(* IEC 61131-3 sources: BODAS-HelloWorld/st/bodas_rc18_12_40/plc_logic/application/02_easyconfig/dsm_easyconfig/structure, 701 files *)

(* ---- dfc_bds_nodeb0x8000-DFC_bds_NoDeb0x8000.st ---- *)
(* --- Interface --- *)
{attribute 'external_name' := 'cmp_rts_DFC_bds_NoDeb0x8000'}
TYPE DFC_bds_NoDeb0x8000 : STRUCT
		DTC            : UDINT := 16#800000;
		DFCid          : UINT  := 721;
		debounceMethod : USINT := NO_DEBOUNCE;
	END_STRUCT
END_TYPE

(* ---- dfc_bds_nodeb0x8001-DFC_bds_NoDeb0x8001.st ---- *)
(* --- Interface --- *)
{attribute 'external_name' := 'cmp_rts_DFC_bds_NoDeb0x8001'}
TYPE DFC_bds_NoDeb0x8001 : STRUCT
		DTC            : UDINT := 16#800100;
		DFCid          : UINT  := 722;
		debounceMethod : USINT := NO_DEBOUNCE;
	END_STRUCT
END_TYPE

(* ---- dfc_bds_nodeb0x8002-DFC_bds_NoDeb0x8002.st ---- *)
(* --- Interface --- *)
{attribute 'external_name' := 'cmp_rts_DFC_bds_NoDeb0x8002'}
TYPE DFC_bds_NoDeb0x8002 : STRUCT
		DTC            : UDINT := 16#800200;
		DFCid          : UINT  := 723;
		debounceMethod : USINT := NO_DEBOUNCE;
	END_STRUCT
END_TYPE

(* ---- dfc_bds_nodeb0x8003-DFC_bds_NoDeb0x8003.st ---- *)
(* --- Interface --- *)
{attribute 'external_name' := 'cmp_rts_DFC_bds_NoDeb0x8003'}
TYPE DFC_bds_NoDeb0x8003 : STRUCT
		DTC            : UDINT := 16#800300;
		DFCid          : UINT  := 724;
		debounceMethod : USINT := NO_DEBOUNCE;
	END_STRUCT
END_TYPE

(* ---- dfc_bds_nodeb0x8004-DFC_bds_NoDeb0x8004.st ---- *)
(* --- Interface --- *)
{attribute 'external_name' := 'cmp_rts_DFC_bds_NoDeb0x8004'}
TYPE DFC_bds_NoDeb0x8004 : STRUCT
		DTC            : UDINT := 16#800400;
		DFCid          : UINT  := 725;
		debounceMethod : USINT := NO_DEBOUNCE;
	END_STRUCT
END_TYPE

(* ---- dfc_bds_nodeb0x8005-DFC_bds_NoDeb0x8005.st ---- *)
(* --- Interface --- *)
{attribute 'external_name' := 'cmp_rts_DFC_bds_NoDeb0x8005'}
TYPE DFC_bds_NoDeb0x8005 : STRUCT
		DTC            : UDINT := 16#800500;
		DFCid          : UINT  := 726;
		debounceMethod : USINT := NO_DEBOUNCE;
	END_STRUCT
END_TYPE

(* ---- dfc_bds_nodeb0x8006-DFC_bds_NoDeb0x8006.st ---- *)
(* --- Interface --- *)
{attribute 'external_name' := 'cmp_rts_DFC_bds_NoDeb0x8006'}
TYPE DFC_bds_NoDeb0x8006 : STRUCT
		DTC            : UDINT := 16#800600;
		DFCid          : UINT  := 727;
		debounceMethod : USINT := NO_DEBOUNCE;
	END_STRUCT
END_TYPE

(* ---- dfc_bds_nodeb0x8007-DFC_bds_NoDeb0x8007.st ---- *)
(* --- Interface --- *)
{attribute 'external_name' := 'cmp_rts_DFC_bds_NoDeb0x8007'}
TYPE DFC_bds_NoDeb0x8007 : STRUCT
		DTC            : UDINT := 16#800700;
		DFCid          : UINT  := 728;
		debounceMethod : USINT := NO_DEBOUNCE;
	END_STRUCT
END_TYPE

(* ---- dfc_bds_nodeb0x8008-DFC_bds_NoDeb0x8008.st ---- *)
(* --- Interface --- *)
{attribute 'external_name' := 'cmp_rts_DFC_bds_NoDeb0x8008'}
TYPE DFC_bds_NoDeb0x8008 : STRUCT
		DTC            : UDINT := 16#800800;
		DFCid          : UINT  := 729;
		debounceMethod : USINT := NO_DEBOUNCE;
	END_STRUCT
END_TYPE

(* ---- dfc_bds_nodeb0x8009-DFC_bds_NoDeb0x8009.st ---- *)
(* --- Interface --- *)
{attribute 'external_name' := 'cmp_rts_DFC_bds_NoDeb0x8009'}
TYPE DFC_bds_NoDeb0x8009 : STRUCT
		DTC            : UDINT := 16#800900;
		DFCid          : UINT  := 730;
		debounceMethod : USINT := NO_DEBOUNCE;
	END_STRUCT
END_TYPE

(* ---- dfc_bds_nodeb0x800a-DFC_bds_NoDeb0x800a.st ---- *)
(* --- Interface --- *)
{attribute 'external_name' := 'cmp_rts_DFC_bds_NoDeb0x800a'}
TYPE DFC_bds_NoDeb0x800a : STRUCT
		DTC            : UDINT := 16#800A00;
		DFCid          : UINT  := 731;
		debounceMethod : USINT := NO_DEBOUNCE;
	END_STRUCT
END_TYPE

(* ---- dfc_bds_nodeb0x800b-DFC_bds_NoDeb0x800b.st ---- *)
(* --- Interface --- *)
{attribute 'external_name' := 'cmp_rts_DFC_bds_NoDeb0x800b'}
TYPE DFC_bds_NoDeb0x800b : STRUCT
		DTC            : UDINT := 16#800B00;
		DFCid          : UINT  := 732;
		debounceMethod : USINT := NO_DEBOUNCE;
	END_STRUCT
END_TYPE

(* ---- dfc_bds_nodeb0x800c-DFC_bds_NoDeb0x800c.st ---- *)
(* --- Interface --- *)
{attribute 'external_name' := 'cmp_rts_DFC_bds_NoDeb0x800c'}
TYPE DFC_bds_NoDeb0x800c : STRUCT
		DTC            : UDINT := 16#800C00;
		DFCid          : UINT  := 733;
		debounceMethod : USINT := NO_DEBOUNCE;
	END_STRUCT
END_TYPE

(* ---- dfc_bds_nodeb0x800d-DFC_bds_NoDeb0x800d.st ---- *)
(* --- Interface --- *)
{attribute 'external_name' := 'cmp_rts_DFC_bds_NoDeb0x800d'}
TYPE DFC_bds_NoDeb0x800d : STRUCT
		DTC            : UDINT := 16#800D00;
		DFCid          : UINT  := 734;
		debounceMethod : USINT := NO_DEBOUNCE;
	END_STRUCT
END_TYPE

(* ---- dfc_bds_nodeb0x800e-DFC_bds_NoDeb0x800e.st ---- *)
(* --- Interface --- *)
{attribute 'external_name' := 'cmp_rts_DFC_bds_NoDeb0x800e'}
TYPE DFC_bds_NoDeb0x800e : STRUCT
		DTC            : UDINT := 16#800E00;
		DFCid          : UINT  := 735;
		debounceMethod : USINT := NO_DEBOUNCE;
	END_STRUCT
END_TYPE

(* ---- dfc_bds_nodeb0x800f-DFC_bds_NoDeb0x800f.st ---- *)
(* --- Interface --- *)
{attribute 'external_name' := 'cmp_rts_DFC_bds_NoDeb0x800f'}
TYPE DFC_bds_NoDeb0x800f : STRUCT
		DTC            : UDINT := 16#800F00;
		DFCid          : UINT  := 736;
		debounceMethod : USINT := NO_DEBOUNCE;
	END_STRUCT
END_TYPE

(* ---- dfc_bds_nodeb0x8010-DFC_bds_NoDeb0x8010.st ---- *)
(* --- Interface --- *)
{attribute 'external_name' := 'cmp_rts_DFC_bds_NoDeb0x8010'}
TYPE DFC_bds_NoDeb0x8010 : STRUCT
		DTC            : UDINT := 16#801000;
		DFCid          : UINT  := 737;
		debounceMethod : USINT := NO_DEBOUNCE;
	END_STRUCT
END_TYPE

(* ---- dfc_bds_nodeb0x8011-DFC_bds_NoDeb0x8011.st ---- *)
(* --- Interface --- *)
{attribute 'external_name' := 'cmp_rts_DFC_bds_NoDeb0x8011'}
TYPE DFC_bds_NoDeb0x8011 : STRUCT
		DTC            : UDINT := 16#801100;
		DFCid          : UINT  := 738;
		debounceMethod : USINT := NO_DEBOUNCE;
	END_STRUCT
END_TYPE

(* ---- dfc_bds_nodeb0x8012-DFC_bds_NoDeb0x8012.st ---- *)
(* --- Interface --- *)
{attribute 'external_name' := 'cmp_rts_DFC_bds_NoDeb0x8012'}
TYPE DFC_bds_NoDeb0x8012 : STRUCT
		DTC            : UDINT := 16#801200;
		DFCid          : UINT  := 739;
		debounceMethod : USINT := NO_DEBOUNCE;
	END_STRUCT
END_TYPE

(* ---- dfc_bds_nodeb0x8013-DFC_bds_NoDeb0x8013.st ---- *)
(* --- Interface --- *)
{attribute 'external_name' := 'cmp_rts_DFC_bds_NoDeb0x8013'}
TYPE DFC_bds_NoDeb0x8013 : STRUCT
		DTC            : UDINT := 16#801300;
		DFCid          : UINT  := 740;
		debounceMethod : USINT := NO_DEBOUNCE;
	END_STRUCT
END_TYPE

(* ---- dfc_bds_nodeb0x8014-DFC_bds_NoDeb0x8014.st ---- *)
(* --- Interface --- *)
{attribute 'external_name' := 'cmp_rts_DFC_bds_NoDeb0x8014'}
TYPE DFC_bds_NoDeb0x8014 : STRUCT
		DTC            : UDINT := 16#801400;
		DFCid          : UINT  := 741;
		debounceMethod : USINT := NO_DEBOUNCE;
	END_STRUCT
END_TYPE

(* ---- dfc_bds_nodeb0x8015-DFC_bds_NoDeb0x8015.st ---- *)
(* --- Interface --- *)
{attribute 'external_name' := 'cmp_rts_DFC_bds_NoDeb0x8015'}
TYPE DFC_bds_NoDeb0x8015 : STRUCT
		DTC            : UDINT := 16#801500;
		DFCid          : UINT  := 742;
		debounceMethod : USINT := NO_DEBOUNCE;
	END_STRUCT
END_TYPE

(* ---- dfc_bds_nodeb0x8016-DFC_bds_NoDeb0x8016.st ---- *)
(* --- Interface --- *)
{attribute 'external_name' := 'cmp_rts_DFC_bds_NoDeb0x8016'}
TYPE DFC_bds_NoDeb0x8016 : STRUCT
		DTC            : UDINT := 16#801600;
		DFCid          : UINT  := 743;
		debounceMethod : USINT := NO_DEBOUNCE;
	END_STRUCT
END_TYPE

(* ---- dfc_bds_nodeb0x8017-DFC_bds_NoDeb0x8017.st ---- *)
(* --- Interface --- *)
{attribute 'external_name' := 'cmp_rts_DFC_bds_NoDeb0x8017'}
TYPE DFC_bds_NoDeb0x8017 : STRUCT
		DTC            : UDINT := 16#801700;
		DFCid          : UINT  := 744;
		debounceMethod : USINT := NO_DEBOUNCE;
	END_STRUCT
END_TYPE

(* ---- dfc_bds_nodeb0x8018-DFC_bds_NoDeb0x8018.st ---- *)
(* --- Interface --- *)
{attribute 'external_name' := 'cmp_rts_DFC_bds_NoDeb0x8018'}
TYPE DFC_bds_NoDeb0x8018 : STRUCT
		DTC            : UDINT := 16#801800;
		DFCid          : UINT  := 745;
		debounceMethod : USINT := NO_DEBOUNCE;
	END_STRUCT
END_TYPE

(* ---- dfc_bds_nodeb0x8019-DFC_bds_NoDeb0x8019.st ---- *)
(* --- Interface --- *)
{attribute 'external_name' := 'cmp_rts_DFC_bds_NoDeb0x8019'}
TYPE DFC_bds_NoDeb0x8019 : STRUCT
		DTC            : UDINT := 16#801900;
		DFCid          : UINT  := 746;
		debounceMethod : USINT := NO_DEBOUNCE;
	END_STRUCT
END_TYPE

(* ---- dfc_bds_nodeb0x801a-DFC_bds_NoDeb0x801a.st ---- *)
(* --- Interface --- *)
{attribute 'external_name' := 'cmp_rts_DFC_bds_NoDeb0x801a'}
TYPE DFC_bds_NoDeb0x801a : STRUCT
		DTC            : UDINT := 16#801A00;
		DFCid          : UINT  := 747;
		debounceMethod : USINT := NO_DEBOUNCE;
	END_STRUCT
END_TYPE

(* ---- dfc_bds_nodeb0x801b-DFC_bds_NoDeb0x801b.st ---- *)
(* --- Interface --- *)
{attribute 'external_name' := 'cmp_rts_DFC_bds_NoDeb0x801b'}
TYPE DFC_bds_NoDeb0x801b : STRUCT
		DTC            : UDINT := 16#801B00;
		DFCid          : UINT  := 748;
		debounceMethod : USINT := NO_DEBOUNCE;
	END_STRUCT
END_TYPE

(* ---- dfc_bds_nodeb0x801c-DFC_bds_NoDeb0x801c.st ---- *)
(* --- Interface --- *)
{attribute 'external_name' := 'cmp_rts_DFC_bds_NoDeb0x801c'}
TYPE DFC_bds_NoDeb0x801c : STRUCT
		DTC            : UDINT := 16#801C00;
		DFCid          : UINT  := 749;
		debounceMethod : USINT := NO_DEBOUNCE;
	END_STRUCT
END_TYPE

(* ---- dfc_bds_nodeb0x801d-DFC_bds_NoDeb0x801d.st ---- *)
(* --- Interface --- *)
{attribute 'external_name' := 'cmp_rts_DFC_bds_NoDeb0x801d'}
TYPE DFC_bds_NoDeb0x801d : STRUCT
		DTC            : UDINT := 16#801D00;
		DFCid          : UINT  := 750;
		debounceMethod : USINT := NO_DEBOUNCE;
	END_STRUCT
END_TYPE

(* ---- dfc_bds_nodeb0x801e-DFC_bds_NoDeb0x801e.st ---- *)
(* --- Interface --- *)
{attribute 'external_name' := 'cmp_rts_DFC_bds_NoDeb0x801e'}
TYPE DFC_bds_NoDeb0x801e : STRUCT
		DTC            : UDINT := 16#801E00;
		DFCid          : UINT  := 751;
		debounceMethod : USINT := NO_DEBOUNCE;
	END_STRUCT
END_TYPE

(* ---- dfc_bds_nodeb0x801f-DFC_bds_NoDeb0x801f.st ---- *)
(* --- Interface --- *)
{attribute 'external_name' := 'cmp_rts_DFC_bds_NoDeb0x801f'}
TYPE DFC_bds_NoDeb0x801f : STRUCT
		DTC            : UDINT := 16#801F00;
		DFCid          : UINT  := 752;
		debounceMethod : USINT := NO_DEBOUNCE;
	END_STRUCT
END_TYPE

(* ---- dfc_bds_nodeb0x8020-DFC_bds_NoDeb0x8020.st ---- *)
(* --- Interface --- *)
{attribute 'external_name' := 'cmp_rts_DFC_bds_NoDeb0x8020'}
TYPE DFC_bds_NoDeb0x8020 : STRUCT
		DTC            : UDINT := 16#802000;
		DFCid          : UINT  := 753;
		debounceMethod : USINT := NO_DEBOUNCE;
	END_STRUCT
END_TYPE

(* ---- dfc_bds_nodeb0x8021-DFC_bds_NoDeb0x8021.st ---- *)
(* --- Interface --- *)
{attribute 'external_name' := 'cmp_rts_DFC_bds_NoDeb0x8021'}
TYPE DFC_bds_NoDeb0x8021 : STRUCT
		DTC            : UDINT := 16#802100;
		DFCid          : UINT  := 754;
		debounceMethod : USINT := NO_DEBOUNCE;
	END_STRUCT
END_TYPE

(* ---- dfc_bds_nodeb0x8022-DFC_bds_NoDeb0x8022.st ---- *)
(* --- Interface --- *)
{attribute 'external_name' := 'cmp_rts_DFC_bds_NoDeb0x8022'}
TYPE DFC_bds_NoDeb0x8022 : STRUCT
		DTC            : UDINT := 16#802200;
		DFCid          : UINT  := 755;
		debounceMethod : USINT := NO_DEBOUNCE;
	END_STRUCT
END_TYPE

(* ---- dfc_bds_nodeb0x8023-DFC_bds_NoDeb0x8023.st ---- *)
(* --- Interface --- *)
{attribute 'external_name' := 'cmp_rts_DFC_bds_NoDeb0x8023'}
TYPE DFC_bds_NoDeb0x8023 : STRUCT
		DTC            : UDINT := 16#802300;
		DFCid          : UINT  := 756;
		debounceMethod : USINT := NO_DEBOUNCE;
	END_STRUCT
END_TYPE

(* ---- dfc_bds_nodeb0x8024-DFC_bds_NoDeb0x8024.st ---- *)
(* --- Interface --- *)
{attribute 'external_name' := 'cmp_rts_DFC_bds_NoDeb0x8024'}
TYPE DFC_bds_NoDeb0x8024 : STRUCT
		DTC            : UDINT := 16#802400;
		DFCid          : UINT  := 757;
		debounceMethod : USINT := NO_DEBOUNCE;
	END_STRUCT
END_TYPE

(* ---- dfc_bds_nodeb0x8025-DFC_bds_NoDeb0x8025.st ---- *)
(* --- Interface --- *)
{attribute 'external_name' := 'cmp_rts_DFC_bds_NoDeb0x8025'}
TYPE DFC_bds_NoDeb0x8025 : STRUCT
		DTC            : UDINT := 16#802500;
		DFCid          : UINT  := 758;
		debounceMethod : USINT := NO_DEBOUNCE;
	END_STRUCT
END_TYPE

(* ---- dfc_bds_nodeb0x8026-DFC_bds_NoDeb0x8026.st ---- *)
(* --- Interface --- *)
{attribute 'external_name' := 'cmp_rts_DFC_bds_NoDeb0x8026'}
TYPE DFC_bds_NoDeb0x8026 : STRUCT
		DTC            : UDINT := 16#802600;
		DFCid          : UINT  := 759;
		debounceMethod : USINT := NO_DEBOUNCE;
	END_STRUCT
END_TYPE

(* ---- dfc_bds_nodeb0x8027-DFC_bds_NoDeb0x8027.st ---- *)
(* --- Interface --- *)
{attribute 'external_name' := 'cmp_rts_DFC_bds_NoDeb0x8027'}
TYPE DFC_bds_NoDeb0x8027 : STRUCT
		DTC            : UDINT := 16#802700;
		DFCid          : UINT  := 760;
		debounceMethod : USINT := NO_DEBOUNCE;
	END_STRUCT
END_TYPE

(* ---- dfc_bds_nodeb0x8028-DFC_bds_NoDeb0x8028.st ---- *)
(* --- Interface --- *)
{attribute 'external_name' := 'cmp_rts_DFC_bds_NoDeb0x8028'}
TYPE DFC_bds_NoDeb0x8028 : STRUCT
		DTC            : UDINT := 16#802800;
		DFCid          : UINT  := 761;
		debounceMethod : USINT := NO_DEBOUNCE;
	END_STRUCT
END_TYPE

(* ---- dfc_bds_nodeb0x8029-DFC_bds_NoDeb0x8029.st ---- *)
(* --- Interface --- *)
{attribute 'external_name' := 'cmp_rts_DFC_bds_NoDeb0x8029'}
TYPE DFC_bds_NoDeb0x8029 : STRUCT
		DTC            : UDINT := 16#802900;
		DFCid          : UINT  := 762;
		debounceMethod : USINT := NO_DEBOUNCE;
	END_STRUCT
END_TYPE

(* ---- dfc_bds_nodeb0x802a-DFC_bds_NoDeb0x802a.st ---- *)
(* --- Interface --- *)
{attribute 'external_name' := 'cmp_rts_DFC_bds_NoDeb0x802a'}
TYPE DFC_bds_NoDeb0x802a : STRUCT
		DTC            : UDINT := 16#802A00;
		DFCid          : UINT  := 763;
		debounceMethod : USINT := NO_DEBOUNCE;
	END_STRUCT
END_TYPE

(* ---- dfc_bds_nodeb0x802b-DFC_bds_NoDeb0x802b.st ---- *)
(* --- Interface --- *)
{attribute 'external_name' := 'cmp_rts_DFC_bds_NoDeb0x802b'}
TYPE DFC_bds_NoDeb0x802b : STRUCT
		DTC            : UDINT := 16#802B00;
		DFCid          : UINT  := 764;
		debounceMethod : USINT := NO_DEBOUNCE;
	END_STRUCT
END_TYPE

(* ---- dfc_bds_nodeb0x802c-DFC_bds_NoDeb0x802c.st ---- *)
(* --- Interface --- *)
{attribute 'external_name' := 'cmp_rts_DFC_bds_NoDeb0x802c'}
TYPE DFC_bds_NoDeb0x802c : STRUCT
		DTC            : UDINT := 16#802C00;
		DFCid          : UINT  := 765;
		debounceMethod : USINT := NO_DEBOUNCE;
	END_STRUCT
END_TYPE

(* ---- dfc_bds_nodeb0x802d-DFC_bds_NoDeb0x802d.st ---- *)
(* --- Interface --- *)
{attribute 'external_name' := 'cmp_rts_DFC_bds_NoDeb0x802d'}
TYPE DFC_bds_NoDeb0x802d : STRUCT
		DTC            : UDINT := 16#802D00;
		DFCid          : UINT  := 766;
		debounceMethod : USINT := NO_DEBOUNCE;
	END_STRUCT
END_TYPE

(* ---- dfc_bds_nodeb0x802e-DFC_bds_NoDeb0x802e.st ---- *)
(* --- Interface --- *)
{attribute 'external_name' := 'cmp_rts_DFC_bds_NoDeb0x802e'}
TYPE DFC_bds_NoDeb0x802e : STRUCT
		DTC            : UDINT := 16#802E00;
		DFCid          : UINT  := 767;
		debounceMethod : USINT := NO_DEBOUNCE;
	END_STRUCT
END_TYPE

(* ---- dfc_bds_nodeb0x802f-DFC_bds_NoDeb0x802f.st ---- *)
(* --- Interface --- *)
{attribute 'external_name' := 'cmp_rts_DFC_bds_NoDeb0x802f'}
TYPE DFC_bds_NoDeb0x802f : STRUCT
		DTC            : UDINT := 16#802F00;
		DFCid          : UINT  := 768;
		debounceMethod : USINT := NO_DEBOUNCE;
	END_STRUCT
END_TYPE

(* ---- dfc_bds_nodeb0x8030-DFC_bds_NoDeb0x8030.st ---- *)
(* --- Interface --- *)
{attribute 'external_name' := 'cmp_rts_DFC_bds_NoDeb0x8030'}
TYPE DFC_bds_NoDeb0x8030 : STRUCT
		DTC            : UDINT := 16#803000;
		DFCid          : UINT  := 769;
		debounceMethod : USINT := NO_DEBOUNCE;
	END_STRUCT
END_TYPE

(* ---- dfc_bds_nodeb0x8031-DFC_bds_NoDeb0x8031.st ---- *)
(* --- Interface --- *)
{attribute 'external_name' := 'cmp_rts_DFC_bds_NoDeb0x8031'}
TYPE DFC_bds_NoDeb0x8031 : STRUCT
		DTC            : UDINT := 16#803100;
		DFCid          : UINT  := 770;
		debounceMethod : USINT := NO_DEBOUNCE;
	END_STRUCT
END_TYPE

(* ---- dfc_bds_nodeb0x8032-DFC_bds_NoDeb0x8032.st ---- *)
(* --- Interface --- *)
{attribute 'external_name' := 'cmp_rts_DFC_bds_NoDeb0x8032'}
TYPE DFC_bds_NoDeb0x8032 : STRUCT
		DTC            : UDINT := 16#803200;
		DFCid          : UINT  := 771;
		debounceMethod : USINT := NO_DEBOUNCE;
	END_STRUCT
END_TYPE

(* ---- dfc_bds_nodeb0x8033-DFC_bds_NoDeb0x8033.st ---- *)
(* --- Interface --- *)
{attribute 'external_name' := 'cmp_rts_DFC_bds_NoDeb0x8033'}
TYPE DFC_bds_NoDeb0x8033 : STRUCT
		DTC            : UDINT := 16#803300;
		DFCid          : UINT  := 772;
		debounceMethod : USINT := NO_DEBOUNCE;
	END_STRUCT
END_TYPE

(* ---- dfc_bds_nodeb0x8034-DFC_bds_NoDeb0x8034.st ---- *)
(* --- Interface --- *)
{attribute 'external_name' := 'cmp_rts_DFC_bds_NoDeb0x8034'}
TYPE DFC_bds_NoDeb0x8034 : STRUCT
		DTC            : UDINT := 16#803400;
		DFCid          : UINT  := 773;
		debounceMethod : USINT := NO_DEBOUNCE;
	END_STRUCT
END_TYPE

(* ---- dfc_bds_nodeb0x8035-DFC_bds_NoDeb0x8035.st ---- *)
(* --- Interface --- *)
{attribute 'external_name' := 'cmp_rts_DFC_bds_NoDeb0x8035'}
TYPE DFC_bds_NoDeb0x8035 : STRUCT
		DTC            : UDINT := 16#803500;
		DFCid          : UINT  := 774;
		debounceMethod : USINT := NO_DEBOUNCE;
	END_STRUCT
END_TYPE

(* ---- dfc_bds_nodeb0x8036-DFC_bds_NoDeb0x8036.st ---- *)
(* --- Interface --- *)
{attribute 'external_name' := 'cmp_rts_DFC_bds_NoDeb0x8036'}
TYPE DFC_bds_NoDeb0x8036 : STRUCT
		DTC            : UDINT := 16#803600;
		DFCid          : UINT  := 775;
		debounceMethod : USINT := NO_DEBOUNCE;
	END_STRUCT
END_TYPE

(* ---- dfc_bds_nodeb0x8037-DFC_bds_NoDeb0x8037.st ---- *)
(* --- Interface --- *)
{attribute 'external_name' := 'cmp_rts_DFC_bds_NoDeb0x8037'}
TYPE DFC_bds_NoDeb0x8037 : STRUCT
		DTC            : UDINT := 16#803700;
		DFCid          : UINT  := 776;
		debounceMethod : USINT := NO_DEBOUNCE;
	END_STRUCT
END_TYPE

(* ---- dfc_bds_nodeb0x8038-DFC_bds_NoDeb0x8038.st ---- *)
(* --- Interface --- *)
{attribute 'external_name' := 'cmp_rts_DFC_bds_NoDeb0x8038'}
TYPE DFC_bds_NoDeb0x8038 : STRUCT
		DTC            : UDINT := 16#803800;
		DFCid          : UINT  := 777;
		debounceMethod : USINT := NO_DEBOUNCE;
	END_STRUCT
END_TYPE

(* ---- dfc_bds_nodeb0x8039-DFC_bds_NoDeb0x8039.st ---- *)
(* --- Interface --- *)
{attribute 'external_name' := 'cmp_rts_DFC_bds_NoDeb0x8039'}
TYPE DFC_bds_NoDeb0x8039 : STRUCT
		DTC            : UDINT := 16#803900;
		DFCid          : UINT  := 778;
		debounceMethod : USINT := NO_DEBOUNCE;
	END_STRUCT
END_TYPE

(* ---- dfc_bds_nodeb0x803a-DFC_bds_NoDeb0x803a.st ---- *)
(* --- Interface --- *)
{attribute 'external_name' := 'cmp_rts_DFC_bds_NoDeb0x803a'}
TYPE DFC_bds_NoDeb0x803a : STRUCT
		DTC            : UDINT := 16#803A00;
		DFCid          : UINT  := 779;
		debounceMethod : USINT := NO_DEBOUNCE;
	END_STRUCT
END_TYPE

(* ---- dfc_bds_nodeb0x803b-DFC_bds_NoDeb0x803b.st ---- *)
(* --- Interface --- *)
{attribute 'external_name' := 'cmp_rts_DFC_bds_NoDeb0x803b'}
TYPE DFC_bds_NoDeb0x803b : STRUCT
		DTC            : UDINT := 16#803B00;
		DFCid          : UINT  := 780;
		debounceMethod : USINT := NO_DEBOUNCE;
	END_STRUCT
END_TYPE

(* ---- dfc_bds_nodeb0x803c-DFC_bds_NoDeb0x803c.st ---- *)
(* --- Interface --- *)
{attribute 'external_name' := 'cmp_rts_DFC_bds_NoDeb0x803c'}
TYPE DFC_bds_NoDeb0x803c : STRUCT
		DTC            : UDINT := 16#803C00;
		DFCid          : UINT  := 781;
		debounceMethod : USINT := NO_DEBOUNCE;
	END_STRUCT
END_TYPE

(* ---- dfc_bds_nodeb0x803d-DFC_bds_NoDeb0x803d.st ---- *)
(* --- Interface --- *)
{attribute 'external_name' := 'cmp_rts_DFC_bds_NoDeb0x803d'}
TYPE DFC_bds_NoDeb0x803d : STRUCT
		DTC            : UDINT := 16#803D00;
		DFCid          : UINT  := 782;
		debounceMethod : USINT := NO_DEBOUNCE;
	END_STRUCT
END_TYPE

(* ---- dfc_bds_nodeb0x803e-DFC_bds_NoDeb0x803e.st ---- *)
(* --- Interface --- *)
{attribute 'external_name' := 'cmp_rts_DFC_bds_NoDeb0x803e'}
TYPE DFC_bds_NoDeb0x803e : STRUCT
		DTC            : UDINT := 16#803E00;
		DFCid          : UINT  := 783;
		debounceMethod : USINT := NO_DEBOUNCE;
	END_STRUCT
END_TYPE

(* ---- dfc_bds_nodeb0x803f-DFC_bds_NoDeb0x803f.st ---- *)
(* --- Interface --- *)
{attribute 'external_name' := 'cmp_rts_DFC_bds_NoDeb0x803f'}
TYPE DFC_bds_NoDeb0x803f : STRUCT
		DTC            : UDINT := 16#803F00;
		DFCid          : UINT  := 784;
		debounceMethod : USINT := NO_DEBOUNCE;
	END_STRUCT
END_TYPE

(* ---- dfc_bds_nodeb0x8040-DFC_bds_NoDeb0x8040.st ---- *)
(* --- Interface --- *)
{attribute 'external_name' := 'cmp_rts_DFC_bds_NoDeb0x8040'}
TYPE DFC_bds_NoDeb0x8040 : STRUCT
		DTC            : UDINT := 16#804000;
		DFCid          : UINT  := 785;
		debounceMethod : USINT := NO_DEBOUNCE;
	END_STRUCT
END_TYPE

(* ---- dfc_bds_nodeb0x8041-DFC_bds_NoDeb0x8041.st ---- *)
(* --- Interface --- *)
{attribute 'external_name' := 'cmp_rts_DFC_bds_NoDeb0x8041'}
TYPE DFC_bds_NoDeb0x8041 : STRUCT
		DTC            : UDINT := 16#804100;
		DFCid          : UINT  := 786;
		debounceMethod : USINT := NO_DEBOUNCE;
	END_STRUCT
END_TYPE

(* ---- dfc_bds_nodeb0x8042-DFC_bds_NoDeb0x8042.st ---- *)
(* --- Interface --- *)
{attribute 'external_name' := 'cmp_rts_DFC_bds_NoDeb0x8042'}
TYPE DFC_bds_NoDeb0x8042 : STRUCT
		DTC            : UDINT := 16#804200;
		DFCid          : UINT  := 787;
		debounceMethod : USINT := NO_DEBOUNCE;
	END_STRUCT
END_TYPE

(* ---- dfc_bds_nodeb0x8043-DFC_bds_NoDeb0x8043.st ---- *)
(* --- Interface --- *)
{attribute 'external_name' := 'cmp_rts_DFC_bds_NoDeb0x8043'}
TYPE DFC_bds_NoDeb0x8043 : STRUCT
		DTC            : UDINT := 16#804300;
		DFCid          : UINT  := 788;
		debounceMethod : USINT := NO_DEBOUNCE;
	END_STRUCT
END_TYPE

(* ---- dfc_bds_nodeb0x8044-DFC_bds_NoDeb0x8044.st ---- *)
(* --- Interface --- *)
{attribute 'external_name' := 'cmp_rts_DFC_bds_NoDeb0x8044'}
TYPE DFC_bds_NoDeb0x8044 : STRUCT
		DTC            : UDINT := 16#804400;
		DFCid          : UINT  := 789;
		debounceMethod : USINT := NO_DEBOUNCE;
	END_STRUCT
END_TYPE

(* ---- dfc_bds_nodeb0x8045-DFC_bds_NoDeb0x8045.st ---- *)
(* --- Interface --- *)
{attribute 'external_name' := 'cmp_rts_DFC_bds_NoDeb0x8045'}
TYPE DFC_bds_NoDeb0x8045 : STRUCT
		DTC            : UDINT := 16#804500;
		DFCid          : UINT  := 790;
		debounceMethod : USINT := NO_DEBOUNCE;
	END_STRUCT
END_TYPE

(* ---- dfc_bds_nodeb0x8046-DFC_bds_NoDeb0x8046.st ---- *)
(* --- Interface --- *)
{attribute 'external_name' := 'cmp_rts_DFC_bds_NoDeb0x8046'}
TYPE DFC_bds_NoDeb0x8046 : STRUCT
		DTC            : UDINT := 16#804600;
		DFCid          : UINT  := 791;
		debounceMethod : USINT := NO_DEBOUNCE;
	END_STRUCT
END_TYPE

(* ---- dfc_bds_nodeb0x8047-DFC_bds_NoDeb0x8047.st ---- *)
(* --- Interface --- *)
{attribute 'external_name' := 'cmp_rts_DFC_bds_NoDeb0x8047'}
TYPE DFC_bds_NoDeb0x8047 : STRUCT
		DTC            : UDINT := 16#804700;
		DFCid          : UINT  := 792;
		debounceMethod : USINT := NO_DEBOUNCE;
	END_STRUCT
END_TYPE

(* ---- dfc_bds_nodeb0x8048-DFC_bds_NoDeb0x8048.st ---- *)
(* --- Interface --- *)
{attribute 'external_name' := 'cmp_rts_DFC_bds_NoDeb0x8048'}
TYPE DFC_bds_NoDeb0x8048 : STRUCT
		DTC            : UDINT := 16#804800;
		DFCid          : UINT  := 793;
		debounceMethod : USINT := NO_DEBOUNCE;
	END_STRUCT
END_TYPE

(* ---- dfc_bds_nodeb0x8049-DFC_bds_NoDeb0x8049.st ---- *)
(* --- Interface --- *)
{attribute 'external_name' := 'cmp_rts_DFC_bds_NoDeb0x8049'}
TYPE DFC_bds_NoDeb0x8049 : STRUCT
		DTC            : UDINT := 16#804900;
		DFCid          : UINT  := 794;
		debounceMethod : USINT := NO_DEBOUNCE;
	END_STRUCT
END_TYPE

(* ---- dfc_bds_nodeb0x804a-DFC_bds_NoDeb0x804a.st ---- *)
(* --- Interface --- *)
{attribute 'external_name' := 'cmp_rts_DFC_bds_NoDeb0x804a'}
TYPE DFC_bds_NoDeb0x804a : STRUCT
		DTC            : UDINT := 16#804A00;
		DFCid          : UINT  := 795;
		debounceMethod : USINT := NO_DEBOUNCE;
	END_STRUCT
END_TYPE

(* ---- dfc_bds_nodeb0x804b-DFC_bds_NoDeb0x804b.st ---- *)
(* --- Interface --- *)
{attribute 'external_name' := 'cmp_rts_DFC_bds_NoDeb0x804b'}
TYPE DFC_bds_NoDeb0x804b : STRUCT
		DTC            : UDINT := 16#804B00;
		DFCid          : UINT  := 796;
		debounceMethod : USINT := NO_DEBOUNCE;
	END_STRUCT
END_TYPE

(* ---- dfc_bds_nodeb0x804c-DFC_bds_NoDeb0x804c.st ---- *)
(* --- Interface --- *)
{attribute 'external_name' := 'cmp_rts_DFC_bds_NoDeb0x804c'}
TYPE DFC_bds_NoDeb0x804c : STRUCT
		DTC            : UDINT := 16#804C00;
		DFCid          : UINT  := 797;
		debounceMethod : USINT := NO_DEBOUNCE;
	END_STRUCT
END_TYPE

(* ---- dfc_bds_nodeb0x804d-DFC_bds_NoDeb0x804d.st ---- *)
(* --- Interface --- *)
{attribute 'external_name' := 'cmp_rts_DFC_bds_NoDeb0x804d'}
TYPE DFC_bds_NoDeb0x804d : STRUCT
		DTC            : UDINT := 16#804D00;
		DFCid          : UINT  := 798;
		debounceMethod : USINT := NO_DEBOUNCE;
	END_STRUCT
END_TYPE

(* ---- dfc_bds_nodeb0x804e-DFC_bds_NoDeb0x804e.st ---- *)
(* --- Interface --- *)
{attribute 'external_name' := 'cmp_rts_DFC_bds_NoDeb0x804e'}
TYPE DFC_bds_NoDeb0x804e : STRUCT
		DTC            : UDINT := 16#804E00;
		DFCid          : UINT  := 799;
		debounceMethod : USINT := NO_DEBOUNCE;
	END_STRUCT
END_TYPE

(* ---- dfc_bds_nodeb0x804f-DFC_bds_NoDeb0x804f.st ---- *)
(* --- Interface --- *)
{attribute 'external_name' := 'cmp_rts_DFC_bds_NoDeb0x804f'}
TYPE DFC_bds_NoDeb0x804f : STRUCT
		DTC            : UDINT := 16#804F00;
		DFCid          : UINT  := 800;
		debounceMethod : USINT := NO_DEBOUNCE;
	END_STRUCT
END_TYPE

(* ---- dfc_bds_nodeb0x8050-DFC_bds_NoDeb0x8050.st ---- *)
(* --- Interface --- *)
{attribute 'external_name' := 'cmp_rts_DFC_bds_NoDeb0x8050'}
TYPE DFC_bds_NoDeb0x8050 : STRUCT
		DTC            : UDINT := 16#805000;
		DFCid          : UINT  := 801;
		debounceMethod : USINT := NO_DEBOUNCE;
	END_STRUCT
END_TYPE

(* ---- dfc_bds_nodeb0x8051-DFC_bds_NoDeb0x8051.st ---- *)
(* --- Interface --- *)
{attribute 'external_name' := 'cmp_rts_DFC_bds_NoDeb0x8051'}
TYPE DFC_bds_NoDeb0x8051 : STRUCT
		DTC            : UDINT := 16#805100;
		DFCid          : UINT  := 802;
		debounceMethod : USINT := NO_DEBOUNCE;
	END_STRUCT
END_TYPE

(* ---- dfc_bds_nodeb0x8052-DFC_bds_NoDeb0x8052.st ---- *)
(* --- Interface --- *)
{attribute 'external_name' := 'cmp_rts_DFC_bds_NoDeb0x8052'}
TYPE DFC_bds_NoDeb0x8052 : STRUCT
		DTC            : UDINT := 16#805200;
		DFCid          : UINT  := 803;
		debounceMethod : USINT := NO_DEBOUNCE;
	END_STRUCT
END_TYPE

(* ---- dfc_bds_nodeb0x8053-DFC_bds_NoDeb0x8053.st ---- *)
(* --- Interface --- *)
{attribute 'external_name' := 'cmp_rts_DFC_bds_NoDeb0x8053'}
TYPE DFC_bds_NoDeb0x8053 : STRUCT
		DTC            : UDINT := 16#805300;
		DFCid          : UINT  := 804;
		debounceMethod : USINT := NO_DEBOUNCE;
	END_STRUCT
END_TYPE

(* ---- dfc_bds_nodeb0x8054-DFC_bds_NoDeb0x8054.st ---- *)
(* --- Interface --- *)
{attribute 'external_name' := 'cmp_rts_DFC_bds_NoDeb0x8054'}
TYPE DFC_bds_NoDeb0x8054 : STRUCT
		DTC            : UDINT := 16#805400;
		DFCid          : UINT  := 805;
		debounceMethod : USINT := NO_DEBOUNCE;
	END_STRUCT
END_TYPE

(* ---- dfc_bds_nodeb0x8055-DFC_bds_NoDeb0x8055.st ---- *)
(* --- Interface --- *)
{attribute 'external_name' := 'cmp_rts_DFC_bds_NoDeb0x8055'}
TYPE DFC_bds_NoDeb0x8055 : STRUCT
		DTC            : UDINT := 16#805500;
		DFCid          : UINT  := 806;
		debounceMethod : USINT := NO_DEBOUNCE;
	END_STRUCT
END_TYPE

(* ---- dfc_bds_nodeb0x8056-DFC_bds_NoDeb0x8056.st ---- *)
(* --- Interface --- *)
{attribute 'external_name' := 'cmp_rts_DFC_bds_NoDeb0x8056'}
TYPE DFC_bds_NoDeb0x8056 : STRUCT
		DTC            : UDINT := 16#805600;
		DFCid          : UINT  := 807;
		debounceMethod : USINT := NO_DEBOUNCE;
	END_STRUCT
END_TYPE

(* ---- dfc_bds_nodeb0x8057-DFC_bds_NoDeb0x8057.st ---- *)
(* --- Interface --- *)
{attribute 'external_name' := 'cmp_rts_DFC_bds_NoDeb0x8057'}
TYPE DFC_bds_NoDeb0x8057 : STRUCT
		DTC            : UDINT := 16#805700;
		DFCid          : UINT  := 808;
		debounceMethod : USINT := NO_DEBOUNCE;
	END_STRUCT
END_TYPE

(* ---- dfc_bds_nodeb0x8058-DFC_bds_NoDeb0x8058.st ---- *)
(* --- Interface --- *)
{attribute 'external_name' := 'cmp_rts_DFC_bds_NoDeb0x8058'}
TYPE DFC_bds_NoDeb0x8058 : STRUCT
		DTC            : UDINT := 16#805800;
		DFCid          : UINT  := 809;
		debounceMethod : USINT := NO_DEBOUNCE;
	END_STRUCT
END_TYPE

(* ---- dfc_bds_nodeb0x8059-DFC_bds_NoDeb0x8059.st ---- *)
(* --- Interface --- *)
{attribute 'external_name' := 'cmp_rts_DFC_bds_NoDeb0x8059'}
TYPE DFC_bds_NoDeb0x8059 : STRUCT
		DTC            : UDINT := 16#805900;
		DFCid          : UINT  := 810;
		debounceMethod : USINT := NO_DEBOUNCE;
	END_STRUCT
END_TYPE

(* ---- dfc_bds_nodeb0x805a-DFC_bds_NoDeb0x805a.st ---- *)
(* --- Interface --- *)
{attribute 'external_name' := 'cmp_rts_DFC_bds_NoDeb0x805a'}
TYPE DFC_bds_NoDeb0x805a : STRUCT
		DTC            : UDINT := 16#805A00;
		DFCid          : UINT  := 811;
		debounceMethod : USINT := NO_DEBOUNCE;
	END_STRUCT
END_TYPE

(* ---- dfc_bds_nodeb0x805b-DFC_bds_NoDeb0x805b.st ---- *)
(* --- Interface --- *)
{attribute 'external_name' := 'cmp_rts_DFC_bds_NoDeb0x805b'}
TYPE DFC_bds_NoDeb0x805b : STRUCT
		DTC            : UDINT := 16#805B00;
		DFCid          : UINT  := 812;
		debounceMethod : USINT := NO_DEBOUNCE;
	END_STRUCT
END_TYPE

(* ---- dfc_bds_nodeb0x805c-DFC_bds_NoDeb0x805c.st ---- *)
(* --- Interface --- *)
{attribute 'external_name' := 'cmp_rts_DFC_bds_NoDeb0x805c'}
TYPE DFC_bds_NoDeb0x805c : STRUCT
		DTC            : UDINT := 16#805C00;
		DFCid          : UINT  := 813;
		debounceMethod : USINT := NO_DEBOUNCE;
	END_STRUCT
END_TYPE

(* ---- dfc_bds_nodeb0x805d-DFC_bds_NoDeb0x805d.st ---- *)
(* --- Interface --- *)
{attribute 'external_name' := 'cmp_rts_DFC_bds_NoDeb0x805d'}
TYPE DFC_bds_NoDeb0x805d : STRUCT
		DTC            : UDINT := 16#805D00;
		DFCid          : UINT  := 814;
		debounceMethod : USINT := NO_DEBOUNCE;
	END_STRUCT
END_TYPE

(* ---- dfc_bds_nodeb0x805e-DFC_bds_NoDeb0x805e.st ---- *)
(* --- Interface --- *)
{attribute 'external_name' := 'cmp_rts_DFC_bds_NoDeb0x805e'}
TYPE DFC_bds_NoDeb0x805e : STRUCT
		DTC            : UDINT := 16#805E00;
		DFCid          : UINT  := 815;
		debounceMethod : USINT := NO_DEBOUNCE;
	END_STRUCT
END_TYPE

(* ---- dfc_bds_nodeb0x805f-DFC_bds_NoDeb0x805f.st ---- *)
(* --- Interface --- *)
{attribute 'external_name' := 'cmp_rts_DFC_bds_NoDeb0x805f'}
TYPE DFC_bds_NoDeb0x805f : STRUCT
		DTC            : UDINT := 16#805F00;
		DFCid          : UINT  := 816;
		debounceMethod : USINT := NO_DEBOUNCE;
	END_STRUCT
END_TYPE

(* ---- dfc_bds_nodeb0x8060-DFC_bds_NoDeb0x8060.st ---- *)
(* --- Interface --- *)
{attribute 'external_name' := 'cmp_rts_DFC_bds_NoDeb0x8060'}
TYPE DFC_bds_NoDeb0x8060 : STRUCT
		DTC            : UDINT := 16#806000;
		DFCid          : UINT  := 817;
		debounceMethod : USINT := NO_DEBOUNCE;
	END_STRUCT
END_TYPE

(* ---- dfc_bds_nodeb0x8061-DFC_bds_NoDeb0x8061.st ---- *)
(* --- Interface --- *)
{attribute 'external_name' := 'cmp_rts_DFC_bds_NoDeb0x8061'}
TYPE DFC_bds_NoDeb0x8061 : STRUCT
		DTC            : UDINT := 16#806100;
		DFCid          : UINT  := 818;
		debounceMethod : USINT := NO_DEBOUNCE;
	END_STRUCT
END_TYPE

(* ---- dfc_bds_nodeb0x8062-DFC_bds_NoDeb0x8062.st ---- *)
(* --- Interface --- *)
{attribute 'external_name' := 'cmp_rts_DFC_bds_NoDeb0x8062'}
TYPE DFC_bds_NoDeb0x8062 : STRUCT
		DTC            : UDINT := 16#806200;
		DFCid          : UINT  := 819;
		debounceMethod : USINT := NO_DEBOUNCE;
	END_STRUCT
END_TYPE

(* ---- dfc_bds_nodeb0x8063-DFC_bds_NoDeb0x8063.st ---- *)
(* --- Interface --- *)
{attribute 'external_name' := 'cmp_rts_DFC_bds_NoDeb0x8063'}
TYPE DFC_bds_NoDeb0x8063 : STRUCT
		DTC            : UDINT := 16#806300;
		DFCid          : UINT  := 106;
		debounceMethod : USINT := TIME_UP_DOWN;
	END_STRUCT
END_TYPE

(* ---- dfc_bds_nodeb0x8064-DFC_bds_NoDeb0x8064.st ---- *)
(* --- Interface --- *)
{attribute 'external_name' := 'cmp_rts_DFC_bds_NoDeb0x8064'}
TYPE DFC_bds_NoDeb0x8064 : STRUCT
		DTC            : UDINT := 16#806400;
		DFCid          : UINT  := 107;
		debounceMethod : USINT := TIME_UP_DOWN;
	END_STRUCT
END_TYPE

(* ---- dfc_bds_nodeb0x8065-DFC_bds_NoDeb0x8065.st ---- *)
(* --- Interface --- *)
{attribute 'external_name' := 'cmp_rts_DFC_bds_NoDeb0x8065'}
TYPE DFC_bds_NoDeb0x8065 : STRUCT
		DTC            : UDINT := 16#806500;
		DFCid          : UINT  := 108;
		debounceMethod : USINT := TIME_UP_DOWN;
	END_STRUCT
END_TYPE

(* ---- dfc_bds_nodeb0x8066-DFC_bds_NoDeb0x8066.st ---- *)
(* --- Interface --- *)
{attribute 'external_name' := 'cmp_rts_DFC_bds_NoDeb0x8066'}
TYPE DFC_bds_NoDeb0x8066 : STRUCT
		DTC            : UDINT := 16#806600;
		DFCid          : UINT  := 109;
		debounceMethod : USINT := TIME_UP_DOWN;
	END_STRUCT
END_TYPE

(* ---- dfc_bds_nodeb0x8067-DFC_bds_NoDeb0x8067.st ---- *)
(* --- Interface --- *)
{attribute 'external_name' := 'cmp_rts_DFC_bds_NoDeb0x8067'}
TYPE DFC_bds_NoDeb0x8067 : STRUCT
		DTC            : UDINT := 16#806700;
		DFCid          : UINT  := 110;
		debounceMethod : USINT := TIME_UP_DOWN;
	END_STRUCT
END_TYPE

(* ---- dfc_bds_nodeb0x8068-DFC_bds_NoDeb0x8068.st ---- *)
(* --- Interface --- *)
{attribute 'external_name' := 'cmp_rts_DFC_bds_NoDeb0x8068'}
TYPE DFC_bds_NoDeb0x8068 : STRUCT
		DTC            : UDINT := 16#806800;
		DFCid          : UINT  := 111;
		debounceMethod : USINT := TIME_UP_DOWN;
	END_STRUCT
END_TYPE

(* ---- dfc_bds_nodeb0x8069-DFC_bds_NoDeb0x8069.st ---- *)
(* --- Interface --- *)
{attribute 'external_name' := 'cmp_rts_DFC_bds_NoDeb0x8069'}
TYPE DFC_bds_NoDeb0x8069 : STRUCT
		DTC            : UDINT := 16#806900;
		DFCid          : UINT  := 112;
		debounceMethod : USINT := TIME_UP_DOWN;
	END_STRUCT
END_TYPE

(* ---- dfc_bds_nodeb0x806a-DFC_bds_NoDeb0x806a.st ---- *)
(* --- Interface --- *)
{attribute 'external_name' := 'cmp_rts_DFC_bds_NoDeb0x806a'}
TYPE DFC_bds_NoDeb0x806a : STRUCT
		DTC            : UDINT := 16#806A00;
		DFCid          : UINT  := 113;
		debounceMethod : USINT := TIME_UP_DOWN;
	END_STRUCT
END_TYPE

(* ---- dfc_bds_nodeb0x806b-DFC_bds_NoDeb0x806b.st ---- *)
(* --- Interface --- *)
{attribute 'external_name' := 'cmp_rts_DFC_bds_NoDeb0x806b'}
TYPE DFC_bds_NoDeb0x806b : STRUCT
		DTC            : UDINT := 16#806B00;
		DFCid          : UINT  := 114;
		debounceMethod : USINT := TIME_UP_DOWN;
	END_STRUCT
END_TYPE

(* ---- dfc_bds_nodeb0x806c-DFC_bds_NoDeb0x806c.st ---- *)
(* --- Interface --- *)
{attribute 'external_name' := 'cmp_rts_DFC_bds_NoDeb0x806c'}
TYPE DFC_bds_NoDeb0x806c : STRUCT
		DTC            : UDINT := 16#806C00;
		DFCid          : UINT  := 115;
		debounceMethod : USINT := TIME_UP_DOWN;
	END_STRUCT
END_TYPE

(* ---- dfc_bds_nodeb0x806d-DFC_bds_NoDeb0x806d.st ---- *)
(* --- Interface --- *)
{attribute 'external_name' := 'cmp_rts_DFC_bds_NoDeb0x806d'}
TYPE DFC_bds_NoDeb0x806d : STRUCT
		DTC            : UDINT := 16#806D00;
		DFCid          : UINT  := 116;
		debounceMethod : USINT := TIME_UP_DOWN;
	END_STRUCT
END_TYPE

(* ---- dfc_bds_nodeb0x806e-DFC_bds_NoDeb0x806e.st ---- *)
(* --- Interface --- *)
{attribute 'external_name' := 'cmp_rts_DFC_bds_NoDeb0x806e'}
TYPE DFC_bds_NoDeb0x806e : STRUCT
		DTC            : UDINT := 16#806E00;
		DFCid          : UINT  := 117;
		debounceMethod : USINT := TIME_UP_DOWN;
	END_STRUCT
END_TYPE

(* ---- dfc_bds_nodeb0x806f-DFC_bds_NoDeb0x806f.st ---- *)
(* --- Interface --- *)
{attribute 'external_name' := 'cmp_rts_DFC_bds_NoDeb0x806f'}
TYPE DFC_bds_NoDeb0x806f : STRUCT
		DTC            : UDINT := 16#806F00;
		DFCid          : UINT  := 118;
		debounceMethod : USINT := TIME_UP_DOWN;
	END_STRUCT
END_TYPE

(* ---- dfc_bds_nodeb0x8070-DFC_bds_NoDeb0x8070.st ---- *)
(* --- Interface --- *)
{attribute 'external_name' := 'cmp_rts_DFC_bds_NoDeb0x8070'}
TYPE DFC_bds_NoDeb0x8070 : STRUCT
		DTC            : UDINT := 16#807000;
		DFCid          : UINT  := 119;
		debounceMethod : USINT := TIME_UP_DOWN;
	END_STRUCT
END_TYPE

(* ---- dfc_bds_nodeb0x8071-DFC_bds_NoDeb0x8071.st ---- *)
(* --- Interface --- *)
{attribute 'external_name' := 'cmp_rts_DFC_bds_NoDeb0x8071'}
TYPE DFC_bds_NoDeb0x8071 : STRUCT
		DTC            : UDINT := 16#807100;
		DFCid          : UINT  := 120;
		debounceMethod : USINT := TIME_UP_DOWN;
	END_STRUCT
END_TYPE

(* ---- dfc_bds_nodeb0x8072-DFC_bds_NoDeb0x8072.st ---- *)
(* --- Interface --- *)
{attribute 'external_name' := 'cmp_rts_DFC_bds_NoDeb0x8072'}
TYPE DFC_bds_NoDeb0x8072 : STRUCT
		DTC            : UDINT := 16#807200;
		DFCid          : UINT  := 121;
		debounceMethod : USINT := TIME_UP_DOWN;
	END_STRUCT
END_TYPE

(* ---- dfc_bds_nodeb0x8073-DFC_bds_NoDeb0x8073.st ---- *)
(* --- Interface --- *)
{attribute 'external_name' := 'cmp_rts_DFC_bds_NoDeb0x8073'}
TYPE DFC_bds_NoDeb0x8073 : STRUCT
		DTC            : UDINT := 16#807300;
		DFCid          : UINT  := 122;
		debounceMethod : USINT := TIME_UP_DOWN;
	END_STRUCT
END_TYPE

(* ---- dfc_bds_nodeb0x8074-DFC_bds_NoDeb0x8074.st ---- *)
(* --- Interface --- *)
{attribute 'external_name' := 'cmp_rts_DFC_bds_NoDeb0x8074'}
TYPE DFC_bds_NoDeb0x8074 : STRUCT
		DTC            : UDINT := 16#807400;
		DFCid          : UINT  := 123;
		debounceMethod : USINT := TIME_UP_DOWN;
	END_STRUCT
END_TYPE

(* ---- dfc_bds_nodeb0x8075-DFC_bds_NoDeb0x8075.st ---- *)
(* --- Interface --- *)
{attribute 'external_name' := 'cmp_rts_DFC_bds_NoDeb0x8075'}
TYPE DFC_bds_NoDeb0x8075 : STRUCT
		DTC            : UDINT := 16#807500;
		DFCid          : UINT  := 124;
		debounceMethod : USINT := TIME_UP_DOWN;
	END_STRUCT
END_TYPE

(* ---- dfc_bds_nodeb0x8076-DFC_bds_NoDeb0x8076.st ---- *)
(* --- Interface --- *)
{attribute 'external_name' := 'cmp_rts_DFC_bds_NoDeb0x8076'}
TYPE DFC_bds_NoDeb0x8076 : STRUCT
		DTC            : UDINT := 16#807600;
		DFCid          : UINT  := 125;
		debounceMethod : USINT := TIME_UP_DOWN;
	END_STRUCT
END_TYPE

(* ---- dfc_bds_nodeb0x8077-DFC_bds_NoDeb0x8077.st ---- *)
(* --- Interface --- *)
{attribute 'external_name' := 'cmp_rts_DFC_bds_NoDeb0x8077'}
TYPE DFC_bds_NoDeb0x8077 : STRUCT
		DTC            : UDINT := 16#807700;
		DFCid          : UINT  := 126;
		debounceMethod : USINT := TIME_UP_DOWN;
	END_STRUCT
END_TYPE

(* ---- dfc_bds_nodeb0x8078-DFC_bds_NoDeb0x8078.st ---- *)
(* --- Interface --- *)
{attribute 'external_name' := 'cmp_rts_DFC_bds_NoDeb0x8078'}
TYPE DFC_bds_NoDeb0x8078 : STRUCT
		DTC            : UDINT := 16#807800;
		DFCid          : UINT  := 127;
		debounceMethod : USINT := TIME_UP_DOWN;
	END_STRUCT
END_TYPE

(* ---- dfc_bds_nodeb0x8079-DFC_bds_NoDeb0x8079.st ---- *)
(* --- Interface --- *)
{attribute 'external_name' := 'cmp_rts_DFC_bds_NoDeb0x8079'}
TYPE DFC_bds_NoDeb0x8079 : STRUCT
		DTC            : UDINT := 16#807900;
		DFCid          : UINT  := 128;
		debounceMethod : USINT := TIME_UP_DOWN;
	END_STRUCT
END_TYPE

(* ---- dfc_bds_nodeb0x807a-DFC_bds_NoDeb0x807a.st ---- *)
(* --- Interface --- *)
{attribute 'external_name' := 'cmp_rts_DFC_bds_NoDeb0x807a'}
TYPE DFC_bds_NoDeb0x807a : STRUCT
		DTC            : UDINT := 16#807A00;
		DFCid          : UINT  := 129;
		debounceMethod : USINT := TIME_UP_DOWN;
	END_STRUCT
END_TYPE

(* ---- dfc_bds_nodeb0x807b-DFC_bds_NoDeb0x807b.st ---- *)
(* --- Interface --- *)
{attribute 'external_name' := 'cmp_rts_DFC_bds_NoDeb0x807b'}
TYPE DFC_bds_NoDeb0x807b : STRUCT
		DTC            : UDINT := 16#807B00;
		DFCid          : UINT  := 130;
		debounceMethod : USINT := TIME_UP_DOWN;
	END_STRUCT
END_TYPE

(* ---- dfc_bds_nodeb0x807c-DFC_bds_NoDeb0x807c.st ---- *)
(* --- Interface --- *)
{attribute 'external_name' := 'cmp_rts_DFC_bds_NoDeb0x807c'}
TYPE DFC_bds_NoDeb0x807c : STRUCT
		DTC            : UDINT := 16#807C00;
		DFCid          : UINT  := 131;
		debounceMethod : USINT := TIME_UP_DOWN;
	END_STRUCT
END_TYPE

(* ---- dfc_bds_nodeb0x807d-DFC_bds_NoDeb0x807d.st ---- *)
(* --- Interface --- *)
{attribute 'external_name' := 'cmp_rts_DFC_bds_NoDeb0x807d'}
TYPE DFC_bds_NoDeb0x807d : STRUCT
		DTC            : UDINT := 16#807D00;
		DFCid          : UINT  := 132;
		debounceMethod : USINT := TIME_UP_DOWN;
	END_STRUCT
END_TYPE

(* ---- dfc_bds_nodeb0x807e-DFC_bds_NoDeb0x807e.st ---- *)
(* --- Interface --- *)
{attribute 'external_name' := 'cmp_rts_DFC_bds_NoDeb0x807e'}
TYPE DFC_bds_NoDeb0x807e : STRUCT
		DTC            : UDINT := 16#807E00;
		DFCid          : UINT  := 133;
		debounceMethod : USINT := TIME_UP_DOWN;
	END_STRUCT
END_TYPE

(* ---- dfc_bds_nodeb0x807f-DFC_bds_NoDeb0x807f.st ---- *)
(* --- Interface --- *)
{attribute 'external_name' := 'cmp_rts_DFC_bds_NoDeb0x807f'}
TYPE DFC_bds_NoDeb0x807f : STRUCT
		DTC            : UDINT := 16#807F00;
		DFCid          : UINT  := 134;
		debounceMethod : USINT := TIME_UP_DOWN;
	END_STRUCT
END_TYPE

(* ---- dfc_bds_nodeb0x8080-DFC_bds_NoDeb0x8080.st ---- *)
(* --- Interface --- *)
{attribute 'external_name' := 'cmp_rts_DFC_bds_NoDeb0x8080'}
TYPE DFC_bds_NoDeb0x8080 : STRUCT
		DTC            : UDINT := 16#808000;
		DFCid          : UINT  := 135;
		debounceMethod : USINT := TIME_UP_DOWN;
	END_STRUCT
END_TYPE

(* ---- dfc_bds_nodeb0x8081-DFC_bds_NoDeb0x8081.st ---- *)
(* --- Interface --- *)
{attribute 'external_name' := 'cmp_rts_DFC_bds_NoDeb0x8081'}
TYPE DFC_bds_NoDeb0x8081 : STRUCT
		DTC            : UDINT := 16#808100;
		DFCid          : UINT  := 136;
		debounceMethod : USINT := TIME_UP_DOWN;
	END_STRUCT
END_TYPE

(* ---- dfc_bds_nodeb0x8082-DFC_bds_NoDeb0x8082.st ---- *)
(* --- Interface --- *)
{attribute 'external_name' := 'cmp_rts_DFC_bds_NoDeb0x8082'}
TYPE DFC_bds_NoDeb0x8082 : STRUCT
		DTC            : UDINT := 16#808200;
		DFCid          : UINT  := 137;
		debounceMethod : USINT := TIME_UP_DOWN;
	END_STRUCT
END_TYPE

(* ---- dfc_bds_nodeb0x8083-DFC_bds_NoDeb0x8083.st ---- *)
(* --- Interface --- *)
{attribute 'external_name' := 'cmp_rts_DFC_bds_NoDeb0x8083'}
TYPE DFC_bds_NoDeb0x8083 : STRUCT
		DTC            : UDINT := 16#808300;
		DFCid          : UINT  := 138;
		debounceMethod : USINT := TIME_UP_DOWN;
	END_STRUCT
END_TYPE

(* ---- dfc_bds_nodeb0x8084-DFC_bds_NoDeb0x8084.st ---- *)
(* --- Interface --- *)
{attribute 'external_name' := 'cmp_rts_DFC_bds_NoDeb0x8084'}
TYPE DFC_bds_NoDeb0x8084 : STRUCT
		DTC            : UDINT := 16#808400;
		DFCid          : UINT  := 139;
		debounceMethod : USINT := TIME_UP_DOWN;
	END_STRUCT
END_TYPE

(* ---- dfc_bds_nodeb0x8085-DFC_bds_NoDeb0x8085.st ---- *)
(* --- Interface --- *)
{attribute 'external_name' := 'cmp_rts_DFC_bds_NoDeb0x8085'}
TYPE DFC_bds_NoDeb0x8085 : STRUCT
		DTC            : UDINT := 16#808500;
		DFCid          : UINT  := 140;
		debounceMethod : USINT := TIME_UP_DOWN;
	END_STRUCT
END_TYPE

(* ---- dfc_bds_nodeb0x8086-DFC_bds_NoDeb0x8086.st ---- *)
(* --- Interface --- *)
{attribute 'external_name' := 'cmp_rts_DFC_bds_NoDeb0x8086'}
TYPE DFC_bds_NoDeb0x8086 : STRUCT
		DTC            : UDINT := 16#808600;
		DFCid          : UINT  := 141;
		debounceMethod : USINT := TIME_UP_DOWN;
	END_STRUCT
END_TYPE

(* ---- dfc_bds_nodeb0x8087-DFC_bds_NoDeb0x8087.st ---- *)
(* --- Interface --- *)
{attribute 'external_name' := 'cmp_rts_DFC_bds_NoDeb0x8087'}
TYPE DFC_bds_NoDeb0x8087 : STRUCT
		DTC            : UDINT := 16#808700;
		DFCid          : UINT  := 142;
		debounceMethod : USINT := TIME_UP_DOWN;
	END_STRUCT
END_TYPE

(* ---- dfc_bds_nodeb0x8088-DFC_bds_NoDeb0x8088.st ---- *)
(* --- Interface --- *)
{attribute 'external_name' := 'cmp_rts_DFC_bds_NoDeb0x8088'}
TYPE DFC_bds_NoDeb0x8088 : STRUCT
		DTC            : UDINT := 16#808800;
		DFCid          : UINT  := 143;
		debounceMethod : USINT := TIME_UP_DOWN;
	END_STRUCT
END_TYPE

(* ---- dfc_bds_nodeb0x8089-DFC_bds_NoDeb0x8089.st ---- *)
(* --- Interface --- *)
{attribute 'external_name' := 'cmp_rts_DFC_bds_NoDeb0x8089'}
TYPE DFC_bds_NoDeb0x8089 : STRUCT
		DTC            : UDINT := 16#808900;
		DFCid          : UINT  := 144;
		debounceMethod : USINT := TIME_UP_DOWN;
	END_STRUCT
END_TYPE

(* ---- dfc_bds_nodeb0x808a-DFC_bds_NoDeb0x808a.st ---- *)
(* --- Interface --- *)
{attribute 'external_name' := 'cmp_rts_DFC_bds_NoDeb0x808a'}
TYPE DFC_bds_NoDeb0x808a : STRUCT
		DTC            : UDINT := 16#808A00;
		DFCid          : UINT  := 145;
		debounceMethod : USINT := TIME_UP_DOWN;
	END_STRUCT
END_TYPE

(* ---- dfc_bds_nodeb0x808b-DFC_bds_NoDeb0x808b.st ---- *)
(* --- Interface --- *)
{attribute 'external_name' := 'cmp_rts_DFC_bds_NoDeb0x808b'}
TYPE DFC_bds_NoDeb0x808b : STRUCT
		DTC            : UDINT := 16#808B00;
		DFCid          : UINT  := 146;
		debounceMethod : USINT := TIME_UP_DOWN;
	END_STRUCT
END_TYPE

(* ---- dfc_bds_nodeb0x808c-DFC_bds_NoDeb0x808c.st ---- *)
(* --- Interface --- *)
{attribute 'external_name' := 'cmp_rts_DFC_bds_NoDeb0x808c'}
TYPE DFC_bds_NoDeb0x808c : STRUCT
		DTC            : UDINT := 16#808C00;
		DFCid          : UINT  := 147;
		debounceMethod : USINT := TIME_UP_DOWN;
	END_STRUCT
END_TYPE

(* ---- dfc_bds_nodeb0x808d-DFC_bds_NoDeb0x808d.st ---- *)
(* --- Interface --- *)
{attribute 'external_name' := 'cmp_rts_DFC_bds_NoDeb0x808d'}
TYPE DFC_bds_NoDeb0x808d : STRUCT
		DTC            : UDINT := 16#808D00;
		DFCid          : UINT  := 148;
		debounceMethod : USINT := TIME_UP_DOWN;
	END_STRUCT
END_TYPE

(* ---- dfc_bds_nodeb0x808e-DFC_bds_NoDeb0x808e.st ---- *)
(* --- Interface --- *)
{attribute 'external_name' := 'cmp_rts_DFC_bds_NoDeb0x808e'}
TYPE DFC_bds_NoDeb0x808e : STRUCT
		DTC            : UDINT := 16#808E00;
		DFCid          : UINT  := 149;
		debounceMethod : USINT := TIME_UP_DOWN;
	END_STRUCT
END_TYPE

(* ---- dfc_bds_nodeb0x808f-DFC_bds_NoDeb0x808f.st ---- *)
(* --- Interface --- *)
{attribute 'external_name' := 'cmp_rts_DFC_bds_NoDeb0x808f'}
TYPE DFC_bds_NoDeb0x808f : STRUCT
		DTC            : UDINT := 16#808F00;
		DFCid          : UINT  := 150;
		debounceMethod : USINT := TIME_UP_DOWN;
	END_STRUCT
END_TYPE

(* ---- dfc_bds_nodeb0x8090-DFC_bds_NoDeb0x8090.st ---- *)
(* --- Interface --- *)
{attribute 'external_name' := 'cmp_rts_DFC_bds_NoDeb0x8090'}
TYPE DFC_bds_NoDeb0x8090 : STRUCT
		DTC            : UDINT := 16#809000;
		DFCid          : UINT  := 151;
		debounceMethod : USINT := TIME_UP_DOWN;
	END_STRUCT
END_TYPE

(* ---- dfc_bds_nodeb0x8091-DFC_bds_NoDeb0x8091.st ---- *)
(* --- Interface --- *)
{attribute 'external_name' := 'cmp_rts_DFC_bds_NoDeb0x8091'}
TYPE DFC_bds_NoDeb0x8091 : STRUCT
		DTC            : UDINT := 16#809100;
		DFCid          : UINT  := 152;
		debounceMethod : USINT := TIME_UP_DOWN;
	END_STRUCT
END_TYPE

(* ---- dfc_bds_nodeb0x8092-DFC_bds_NoDeb0x8092.st ---- *)
(* --- Interface --- *)
{attribute 'external_name' := 'cmp_rts_DFC_bds_NoDeb0x8092'}
TYPE DFC_bds_NoDeb0x8092 : STRUCT
		DTC            : UDINT := 16#809200;
		DFCid          : UINT  := 153;
		debounceMethod : USINT := TIME_UP_DOWN;
	END_STRUCT
END_TYPE

(* ---- dfc_bds_nodeb0x8093-DFC_bds_NoDeb0x8093.st ---- *)
(* --- Interface --- *)
{attribute 'external_name' := 'cmp_rts_DFC_bds_NoDeb0x8093'}
TYPE DFC_bds_NoDeb0x8093 : STRUCT
		DTC            : UDINT := 16#809300;
		DFCid          : UINT  := 154;
		debounceMethod : USINT := TIME_UP_DOWN;
	END_STRUCT
END_TYPE

(* ---- dfc_bds_nodeb0x8094-DFC_bds_NoDeb0x8094.st ---- *)
(* --- Interface --- *)
{attribute 'external_name' := 'cmp_rts_DFC_bds_NoDeb0x8094'}
TYPE DFC_bds_NoDeb0x8094 : STRUCT
		DTC            : UDINT := 16#809400;
		DFCid          : UINT  := 155;
		debounceMethod : USINT := TIME_UP_DOWN;
	END_STRUCT
END_TYPE

(* ---- dfc_bds_nodeb0x8095-DFC_bds_NoDeb0x8095.st ---- *)
(* --- Interface --- *)
{attribute 'external_name' := 'cmp_rts_DFC_bds_NoDeb0x8095'}
TYPE DFC_bds_NoDeb0x8095 : STRUCT
		DTC            : UDINT := 16#809500;
		DFCid          : UINT  := 156;
		debounceMethod : USINT := TIME_UP_DOWN;
	END_STRUCT
END_TYPE

(* ---- dfc_bds_nodeb0x8096-DFC_bds_NoDeb0x8096.st ---- *)
(* --- Interface --- *)
{attribute 'external_name' := 'cmp_rts_DFC_bds_NoDeb0x8096'}
TYPE DFC_bds_NoDeb0x8096 : STRUCT
		DTC            : UDINT := 16#809600;
		DFCid          : UINT  := 157;
		debounceMethod : USINT := TIME_UP_DOWN;
	END_STRUCT
END_TYPE

(* ---- dfc_bds_nodeb0x8097-DFC_bds_NoDeb0x8097.st ---- *)
(* --- Interface --- *)
{attribute 'external_name' := 'cmp_rts_DFC_bds_NoDeb0x8097'}
TYPE DFC_bds_NoDeb0x8097 : STRUCT
		DTC            : UDINT := 16#809700;
		DFCid          : UINT  := 158;
		debounceMethod : USINT := TIME_UP_DOWN;
	END_STRUCT
END_TYPE

(* ---- dfc_bds_nodeb0x8098-DFC_bds_NoDeb0x8098.st ---- *)
(* --- Interface --- *)
{attribute 'external_name' := 'cmp_rts_DFC_bds_NoDeb0x8098'}
TYPE DFC_bds_NoDeb0x8098 : STRUCT
		DTC            : UDINT := 16#809800;
		DFCid          : UINT  := 159;
		debounceMethod : USINT := TIME_UP_DOWN;
	END_STRUCT
END_TYPE

(* ---- dfc_bds_nodeb0x8099-DFC_bds_NoDeb0x8099.st ---- *)
(* --- Interface --- *)
{attribute 'external_name' := 'cmp_rts_DFC_bds_NoDeb0x8099'}
TYPE DFC_bds_NoDeb0x8099 : STRUCT
		DTC            : UDINT := 16#809900;
		DFCid          : UINT  := 160;
		debounceMethod : USINT := TIME_UP_DOWN;
	END_STRUCT
END_TYPE

(* ---- dfc_bds_nodeb0x809a-DFC_bds_NoDeb0x809a.st ---- *)
(* --- Interface --- *)
{attribute 'external_name' := 'cmp_rts_DFC_bds_NoDeb0x809a'}
TYPE DFC_bds_NoDeb0x809a : STRUCT
		DTC            : UDINT := 16#809A00;
		DFCid          : UINT  := 161;
		debounceMethod : USINT := TIME_UP_DOWN;
	END_STRUCT
END_TYPE

(* ---- dfc_bds_nodeb0x809b-DFC_bds_NoDeb0x809b.st ---- *)
(* --- Interface --- *)
{attribute 'external_name' := 'cmp_rts_DFC_bds_NoDeb0x809b'}
TYPE DFC_bds_NoDeb0x809b : STRUCT
		DTC            : UDINT := 16#809B00;
		DFCid          : UINT  := 162;
		debounceMethod : USINT := TIME_UP_DOWN;
	END_STRUCT
END_TYPE

(* ---- dfc_bds_nodeb0x809c-DFC_bds_NoDeb0x809c.st ---- *)
(* --- Interface --- *)
{attribute 'external_name' := 'cmp_rts_DFC_bds_NoDeb0x809c'}
TYPE DFC_bds_NoDeb0x809c : STRUCT
		DTC            : UDINT := 16#809C00;
		DFCid          : UINT  := 163;
		debounceMethod : USINT := TIME_UP_DOWN;
	END_STRUCT
END_TYPE

(* ---- dfc_bds_nodeb0x809d-DFC_bds_NoDeb0x809d.st ---- *)
(* --- Interface --- *)
{attribute 'external_name' := 'cmp_rts_DFC_bds_NoDeb0x809d'}
TYPE DFC_bds_NoDeb0x809d : STRUCT
		DTC            : UDINT := 16#809D00;
		DFCid          : UINT  := 164;
		debounceMethod : USINT := TIME_UP_DOWN;
	END_STRUCT
END_TYPE

(* ---- dfc_bds_nodeb0x809e-DFC_bds_NoDeb0x809e.st ---- *)
(* --- Interface --- *)
{attribute 'external_name' := 'cmp_rts_DFC_bds_NoDeb0x809e'}
TYPE DFC_bds_NoDeb0x809e : STRUCT
		DTC            : UDINT := 16#809E00;
		DFCid          : UINT  := 165;
		debounceMethod : USINT := TIME_UP_DOWN;
	END_STRUCT
END_TYPE

(* ---- dfc_bds_nodeb0x809f-DFC_bds_NoDeb0x809f.st ---- *)
(* --- Interface --- *)
{attribute 'external_name' := 'cmp_rts_DFC_bds_NoDeb0x809f'}
TYPE DFC_bds_NoDeb0x809f : STRUCT
		DTC            : UDINT := 16#809F00;
		DFCid          : UINT  := 166;
		debounceMethod : USINT := TIME_UP_DOWN;
	END_STRUCT
END_TYPE

(* ---- dfc_bds_nodeb0x80a0-DFC_bds_NoDeb0x80a0.st ---- *)
(* --- Interface --- *)
{attribute 'external_name' := 'cmp_rts_DFC_bds_NoDeb0x80a0'}
TYPE DFC_bds_NoDeb0x80a0 : STRUCT
		DTC            : UDINT := 16#80A000;
		DFCid          : UINT  := 167;
		debounceMethod : USINT := TIME_UP_DOWN;
	END_STRUCT
END_TYPE

(* ---- dfc_bds_nodeb0x80a1-DFC_bds_NoDeb0x80a1.st ---- *)
(* --- Interface --- *)
{attribute 'external_name' := 'cmp_rts_DFC_bds_NoDeb0x80a1'}
TYPE DFC_bds_NoDeb0x80a1 : STRUCT
		DTC            : UDINT := 16#80A100;
		DFCid          : UINT  := 168;
		debounceMethod : USINT := TIME_UP_DOWN;
	END_STRUCT
END_TYPE

(* ---- dfc_bds_nodeb0x80a2-DFC_bds_NoDeb0x80a2.st ---- *)
(* --- Interface --- *)
{attribute 'external_name' := 'cmp_rts_DFC_bds_NoDeb0x80a2'}
TYPE DFC_bds_NoDeb0x80a2 : STRUCT
		DTC            : UDINT := 16#80A200;
		DFCid          : UINT  := 169;
		debounceMethod : USINT := TIME_UP_DOWN;
	END_STRUCT
END_TYPE

(* ---- dfc_bds_nodeb0x80a3-DFC_bds_NoDeb0x80a3.st ---- *)
(* --- Interface --- *)
{attribute 'external_name' := 'cmp_rts_DFC_bds_NoDeb0x80a3'}
TYPE DFC_bds_NoDeb0x80a3 : STRUCT
		DTC            : UDINT := 16#80A300;
		DFCid          : UINT  := 170;
		debounceMethod : USINT := TIME_UP_DOWN;
	END_STRUCT
END_TYPE

(* ---- dfc_bds_nodeb0x80a4-DFC_bds_NoDeb0x80a4.st ---- *)
(* --- Interface --- *)
{attribute 'external_name' := 'cmp_rts_DFC_bds_NoDeb0x80a4'}
TYPE DFC_bds_NoDeb0x80a4 : STRUCT
		DTC            : UDINT := 16#80A400;
		DFCid          : UINT  := 171;
		debounceMethod : USINT := TIME_UP_DOWN;
	END_STRUCT
END_TYPE

(* ---- dfc_bds_nodeb0x80a5-DFC_bds_NoDeb0x80a5.st ---- *)
(* --- Interface --- *)
{attribute 'external_name' := 'cmp_rts_DFC_bds_NoDeb0x80a5'}
TYPE DFC_bds_NoDeb0x80a5 : STRUCT
		DTC            : UDINT := 16#80A500;
		DFCid          : UINT  := 172;
		debounceMethod : USINT := TIME_UP_DOWN;
	END_STRUCT
END_TYPE

(* ---- dfc_bds_nodeb0x80a6-DFC_bds_NoDeb0x80a6.st ---- *)
(* --- Interface --- *)
{attribute 'external_name' := 'cmp_rts_DFC_bds_NoDeb0x80a6'}
TYPE DFC_bds_NoDeb0x80a6 : STRUCT
		DTC            : UDINT := 16#80A600;
		DFCid          : UINT  := 173;
		debounceMethod : USINT := TIME_UP_DOWN;
	END_STRUCT
END_TYPE

(* ---- dfc_bds_nodeb0x80a7-DFC_bds_NoDeb0x80a7.st ---- *)
(* --- Interface --- *)
{attribute 'external_name' := 'cmp_rts_DFC_bds_NoDeb0x80a7'}
TYPE DFC_bds_NoDeb0x80a7 : STRUCT
		DTC            : UDINT := 16#80A700;
		DFCid          : UINT  := 174;
		debounceMethod : USINT := TIME_UP_DOWN;
	END_STRUCT
END_TYPE

(* ---- dfc_bds_nodeb0x80a8-DFC_bds_NoDeb0x80a8.st ---- *)
(* --- Interface --- *)
{attribute 'external_name' := 'cmp_rts_DFC_bds_NoDeb0x80a8'}
TYPE DFC_bds_NoDeb0x80a8 : STRUCT
		DTC            : UDINT := 16#80A800;
		DFCid          : UINT  := 175;
		debounceMethod : USINT := TIME_UP_DOWN;
	END_STRUCT
END_TYPE

(* ---- dfc_bds_nodeb0x80a9-DFC_bds_NoDeb0x80a9.st ---- *)
(* --- Interface --- *)
{attribute 'external_name' := 'cmp_rts_DFC_bds_NoDeb0x80a9'}
TYPE DFC_bds_NoDeb0x80a9 : STRUCT
		DTC            : UDINT := 16#80A900;
		DFCid          : UINT  := 176;
		debounceMethod : USINT := TIME_UP_DOWN;
	END_STRUCT
END_TYPE

(* ---- dfc_bds_nodeb0x80aa-DFC_bds_NoDeb0x80aa.st ---- *)
(* --- Interface --- *)
{attribute 'external_name' := 'cmp_rts_DFC_bds_NoDeb0x80aa'}
TYPE DFC_bds_NoDeb0x80aa : STRUCT
		DTC            : UDINT := 16#80AA00;
		DFCid          : UINT  := 177;
		debounceMethod : USINT := TIME_UP_DOWN;
	END_STRUCT
END_TYPE

(* ---- dfc_bds_nodeb0x80ab-DFC_bds_NoDeb0x80ab.st ---- *)
(* --- Interface --- *)
{attribute 'external_name' := 'cmp_rts_DFC_bds_NoDeb0x80ab'}
TYPE DFC_bds_NoDeb0x80ab : STRUCT
		DTC            : UDINT := 16#80AB00;
		DFCid          : UINT  := 178;
		debounceMethod : USINT := TIME_UP_DOWN;
	END_STRUCT
END_TYPE

(* ---- dfc_bds_nodeb0x80ac-DFC_bds_NoDeb0x80ac.st ---- *)
(* --- Interface --- *)
{attribute 'external_name' := 'cmp_rts_DFC_bds_NoDeb0x80ac'}
TYPE DFC_bds_NoDeb0x80ac : STRUCT
		DTC            : UDINT := 16#80AC00;
		DFCid          : UINT  := 179;
		debounceMethod : USINT := TIME_UP_DOWN;
	END_STRUCT
END_TYPE

(* ---- dfc_bds_nodeb0x80ad-DFC_bds_NoDeb0x80ad.st ---- *)
(* --- Interface --- *)
{attribute 'external_name' := 'cmp_rts_DFC_bds_NoDeb0x80ad'}
TYPE DFC_bds_NoDeb0x80ad : STRUCT
		DTC            : UDINT := 16#80AD00;
		DFCid          : UINT  := 180;
		debounceMethod : USINT := TIME_UP_DOWN;
	END_STRUCT
END_TYPE

(* ---- dfc_bds_nodeb0x80ae-DFC_bds_NoDeb0x80ae.st ---- *)
(* --- Interface --- *)
{attribute 'external_name' := 'cmp_rts_DFC_bds_NoDeb0x80ae'}
TYPE DFC_bds_NoDeb0x80ae : STRUCT
		DTC            : UDINT := 16#80AE00;
		DFCid          : UINT  := 181;
		debounceMethod : USINT := TIME_UP_DOWN;
	END_STRUCT
END_TYPE

(* ---- dfc_bds_nodeb0x80af-DFC_bds_NoDeb0x80af.st ---- *)
(* --- Interface --- *)
{attribute 'external_name' := 'cmp_rts_DFC_bds_NoDeb0x80af'}
TYPE DFC_bds_NoDeb0x80af : STRUCT
		DTC            : UDINT := 16#80AF00;
		DFCid          : UINT  := 182;
		debounceMethod : USINT := TIME_UP_DOWN;
	END_STRUCT
END_TYPE

(* ---- dfc_bds_nodeb0x80b0-DFC_bds_NoDeb0x80b0.st ---- *)
(* --- Interface --- *)
{attribute 'external_name' := 'cmp_rts_DFC_bds_NoDeb0x80b0'}
TYPE DFC_bds_NoDeb0x80b0 : STRUCT
		DTC            : UDINT := 16#80B000;
		DFCid          : UINT  := 183;
		debounceMethod : USINT := TIME_UP_DOWN;
	END_STRUCT
END_TYPE

(* ---- dfc_bds_nodeb0x80b1-DFC_bds_NoDeb0x80b1.st ---- *)
(* --- Interface --- *)
{attribute 'external_name' := 'cmp_rts_DFC_bds_NoDeb0x80b1'}
TYPE DFC_bds_NoDeb0x80b1 : STRUCT
		DTC            : UDINT := 16#80B100;
		DFCid          : UINT  := 184;
		debounceMethod : USINT := TIME_UP_DOWN;
	END_STRUCT
END_TYPE

(* ---- dfc_bds_nodeb0x80b2-DFC_bds_NoDeb0x80b2.st ---- *)
(* --- Interface --- *)
{attribute 'external_name' := 'cmp_rts_DFC_bds_NoDeb0x80b2'}
TYPE DFC_bds_NoDeb0x80b2 : STRUCT
		DTC            : UDINT := 16#80B200;
		DFCid          : UINT  := 185;
		debounceMethod : USINT := TIME_UP_DOWN;
	END_STRUCT
END_TYPE

(* ---- dfc_bds_nodeb0x80b3-DFC_bds_NoDeb0x80b3.st ---- *)
(* --- Interface --- *)
{attribute 'external_name' := 'cmp_rts_DFC_bds_NoDeb0x80b3'}
TYPE DFC_bds_NoDeb0x80b3 : STRUCT
		DTC            : UDINT := 16#80B300;
		DFCid          : UINT  := 186;
		debounceMethod : USINT := TIME_UP_DOWN;
	END_STRUCT
END_TYPE

(* ---- dfc_bds_nodeb0x80b4-DFC_bds_NoDeb0x80b4.st ---- *)
(* --- Interface --- *)
{attribute 'external_name' := 'cmp_rts_DFC_bds_NoDeb0x80b4'}
TYPE DFC_bds_NoDeb0x80b4 : STRUCT
		DTC            : UDINT := 16#80B400;
		DFCid          : UINT  := 187;
		debounceMethod : USINT := TIME_UP_DOWN;
	END_STRUCT
END_TYPE

(* ---- dfc_bds_nodeb0x80b5-DFC_bds_NoDeb0x80b5.st ---- *)
(* --- Interface --- *)
{attribute 'external_name' := 'cmp_rts_DFC_bds_NoDeb0x80b5'}
TYPE DFC_bds_NoDeb0x80b5 : STRUCT
		DTC            : UDINT := 16#80B500;
		DFCid          : UINT  := 188;
		debounceMethod : USINT := TIME_UP_DOWN;
	END_STRUCT
END_TYPE

(* ---- dfc_bds_nodeb0x80b6-DFC_bds_NoDeb0x80b6.st ---- *)
(* --- Interface --- *)
{attribute 'external_name' := 'cmp_rts_DFC_bds_NoDeb0x80b6'}
TYPE DFC_bds_NoDeb0x80b6 : STRUCT
		DTC            : UDINT := 16#80B600;
		DFCid          : UINT  := 189;
		debounceMethod : USINT := TIME_UP_DOWN;
	END_STRUCT
END_TYPE

(* ---- dfc_bds_nodeb0x80b7-DFC_bds_NoDeb0x80b7.st ---- *)
(* --- Interface --- *)
{attribute 'external_name' := 'cmp_rts_DFC_bds_NoDeb0x80b7'}
TYPE DFC_bds_NoDeb0x80b7 : STRUCT
		DTC            : UDINT := 16#80B700;
		DFCid          : UINT  := 190;
		debounceMethod : USINT := TIME_UP_DOWN;
	END_STRUCT
END_TYPE

(* ---- dfc_bds_nodeb0x80b8-DFC_bds_NoDeb0x80b8.st ---- *)
(* --- Interface --- *)
{attribute 'external_name' := 'cmp_rts_DFC_bds_NoDeb0x80b8'}
TYPE DFC_bds_NoDeb0x80b8 : STRUCT
		DTC            : UDINT := 16#80B800;
		DFCid          : UINT  := 191;
		debounceMethod : USINT := TIME_UP_DOWN;
	END_STRUCT
END_TYPE

(* ---- dfc_bds_nodeb0x80b9-DFC_bds_NoDeb0x80b9.st ---- *)
(* --- Interface --- *)
{attribute 'external_name' := 'cmp_rts_DFC_bds_NoDeb0x80b9'}
TYPE DFC_bds_NoDeb0x80b9 : STRUCT
		DTC            : UDINT := 16#80B900;
		DFCid          : UINT  := 192;
		debounceMethod : USINT := TIME_UP_DOWN;
	END_STRUCT
END_TYPE

(* ---- dfc_bds_nodeb0x80ba-DFC_bds_NoDeb0x80ba.st ---- *)
(* --- Interface --- *)
{attribute 'external_name' := 'cmp_rts_DFC_bds_NoDeb0x80ba'}
TYPE DFC_bds_NoDeb0x80ba : STRUCT
		DTC            : UDINT := 16#80BA00;
		DFCid          : UINT  := 193;
		debounceMethod : USINT := TIME_UP_DOWN;
	END_STRUCT
END_TYPE

(* ---- dfc_bds_nodeb0x80bb-DFC_bds_NoDeb0x80bb.st ---- *)
(* --- Interface --- *)
{attribute 'external_name' := 'cmp_rts_DFC_bds_NoDeb0x80bb'}
TYPE DFC_bds_NoDeb0x80bb : STRUCT
		DTC            : UDINT := 16#80BB00;
		DFCid          : UINT  := 194;
		debounceMethod : USINT := TIME_UP_DOWN;
	END_STRUCT
END_TYPE

(* ---- dfc_bds_nodeb0x80bc-DFC_bds_NoDeb0x80bc.st ---- *)
(* --- Interface --- *)
{attribute 'external_name' := 'cmp_rts_DFC_bds_NoDeb0x80bc'}
TYPE DFC_bds_NoDeb0x80bc : STRUCT
		DTC            : UDINT := 16#80BC00;
		DFCid          : UINT  := 195;
		debounceMethod : USINT := TIME_UP_DOWN;
	END_STRUCT
END_TYPE

(* ---- dfc_bds_nodeb0x80bd-DFC_bds_NoDeb0x80bd.st ---- *)
(* --- Interface --- *)
{attribute 'external_name' := 'cmp_rts_DFC_bds_NoDeb0x80bd'}
TYPE DFC_bds_NoDeb0x80bd : STRUCT
		DTC            : UDINT := 16#80BD00;
		DFCid          : UINT  := 196;
		debounceMethod : USINT := TIME_UP_DOWN;
	END_STRUCT
END_TYPE

(* ---- dfc_bds_nodeb0x80be-DFC_bds_NoDeb0x80be.st ---- *)
(* --- Interface --- *)
{attribute 'external_name' := 'cmp_rts_DFC_bds_NoDeb0x80be'}
TYPE DFC_bds_NoDeb0x80be : STRUCT
		DTC            : UDINT := 16#80BE00;
		DFCid          : UINT  := 197;
		debounceMethod : USINT := TIME_UP_DOWN;
	END_STRUCT
END_TYPE

(* ---- dfc_bds_nodeb0x80bf-DFC_bds_NoDeb0x80bf.st ---- *)
(* --- Interface --- *)
{attribute 'external_name' := 'cmp_rts_DFC_bds_NoDeb0x80bf'}
TYPE DFC_bds_NoDeb0x80bf : STRUCT
		DTC            : UDINT := 16#80BF00;
		DFCid          : UINT  := 198;
		debounceMethod : USINT := TIME_UP_DOWN;
	END_STRUCT
END_TYPE

(* ---- dfc_bds_nodeb0x80c0-DFC_bds_NoDeb0x80c0.st ---- *)
(* --- Interface --- *)
{attribute 'external_name' := 'cmp_rts_DFC_bds_NoDeb0x80c0'}
TYPE DFC_bds_NoDeb0x80c0 : STRUCT
		DTC            : UDINT := 16#80C000;
		DFCid          : UINT  := 199;
		debounceMethod : USINT := TIME_UP_DOWN;
	END_STRUCT
END_TYPE

(* ---- dfc_bds_nodeb0x80c1-DFC_bds_NoDeb0x80c1.st ---- *)
(* --- Interface --- *)
{attribute 'external_name' := 'cmp_rts_DFC_bds_NoDeb0x80c1'}
TYPE DFC_bds_NoDeb0x80c1 : STRUCT
		DTC            : UDINT := 16#80C100;
		DFCid          : UINT  := 200;
		debounceMethod : USINT := TIME_UP_DOWN;
	END_STRUCT
END_TYPE

(* ---- dfc_bds_nodeb0x80c2-DFC_bds_NoDeb0x80c2.st ---- *)
(* --- Interface --- *)
{attribute 'external_name' := 'cmp_rts_DFC_bds_NoDeb0x80c2'}
TYPE DFC_bds_NoDeb0x80c2 : STRUCT
		DTC            : UDINT := 16#80C200;
		DFCid          : UINT  := 201;
		debounceMethod : USINT := TIME_UP_DOWN;
	END_STRUCT
END_TYPE

(* ---- dfc_bds_nodeb0x80c3-DFC_bds_NoDeb0x80c3.st ---- *)
(* --- Interface --- *)
{attribute 'external_name' := 'cmp_rts_DFC_bds_NoDeb0x80c3'}
TYPE DFC_bds_NoDeb0x80c3 : STRUCT
		DTC            : UDINT := 16#80C300;
		DFCid          : UINT  := 202;
		debounceMethod : USINT := TIME_UP_DOWN;
	END_STRUCT
END_TYPE

(* ---- dfc_bds_nodeb0x80c4-DFC_bds_NoDeb0x80c4.st ---- *)
(* --- Interface --- *)
{attribute 'external_name' := 'cmp_rts_DFC_bds_NoDeb0x80c4'}
TYPE DFC_bds_NoDeb0x80c4 : STRUCT
		DTC            : UDINT := 16#80C400;
		DFCid          : UINT  := 203;
		debounceMethod : USINT := TIME_UP_DOWN;
	END_STRUCT
END_TYPE

(* ---- dfc_bds_nodeb0x80c5-DFC_bds_NoDeb0x80c5.st ---- *)
(* --- Interface --- *)
{attribute 'external_name' := 'cmp_rts_DFC_bds_NoDeb0x80c5'}
TYPE DFC_bds_NoDeb0x80c5 : STRUCT
		DTC            : UDINT := 16#80C500;
		DFCid          : UINT  := 204;
		debounceMethod : USINT := TIME_UP_DOWN;
	END_STRUCT
END_TYPE

(* ---- dfc_bds_nodeb0x80c6-DFC_bds_NoDeb0x80c6.st ---- *)
(* --- Interface --- *)
{attribute 'external_name' := 'cmp_rts_DFC_bds_NoDeb0x80c6'}
TYPE DFC_bds_NoDeb0x80c6 : STRUCT
		DTC            : UDINT := 16#80C600;
		DFCid          : UINT  := 205;
		debounceMethod : USINT := TIME_UP_DOWN;
	END_STRUCT
END_TYPE

(* ---- dfc_bds_nodeb0x80c7-DFC_bds_NoDeb0x80c7.st ---- *)
(* --- Interface --- *)
{attribute 'external_name' := 'cmp_rts_DFC_bds_NoDeb0x80c7'}
TYPE DFC_bds_NoDeb0x80c7 : STRUCT
		DTC            : UDINT := 16#80C700;
		DFCid          : UINT  := 1;
		debounceMethod : USINT := TIME_IN_ROW;
	END_STRUCT
END_TYPE

(* ---- dfc_bds_nodeb0x80c8-DFC_bds_NoDeb0x80c8.st ---- *)
(* --- Interface --- *)
{attribute 'external_name' := 'cmp_rts_DFC_bds_NoDeb0x80c8'}
TYPE DFC_bds_NoDeb0x80c8 : STRUCT
		DTC            : UDINT := 16#80C800;
		DFCid          : UINT  := 2;
		debounceMethod : USINT := TIME_IN_ROW;
	END_STRUCT
END_TYPE

(* ---- dfc_bds_nodeb0x80c9-DFC_bds_NoDeb0x80c9.st ---- *)
(* --- Interface --- *)
{attribute 'external_name' := 'cmp_rts_DFC_bds_NoDeb0x80c9'}
TYPE DFC_bds_NoDeb0x80c9 : STRUCT
		DTC            : UDINT := 16#80C900;
		DFCid          : UINT  := 3;
		debounceMethod : USINT := TIME_IN_ROW;
	END_STRUCT
END_TYPE

(* ---- dfc_bds_nodeb0x80ca-DFC_bds_NoDeb0x80ca.st ---- *)
(* --- Interface --- *)
{attribute 'external_name' := 'cmp_rts_DFC_bds_NoDeb0x80ca'}
TYPE DFC_bds_NoDeb0x80ca : STRUCT
		DTC            : UDINT := 16#80CA00;
		DFCid          : UINT  := 4;
		debounceMethod : USINT := TIME_IN_ROW;
	END_STRUCT
END_TYPE

(* ---- dfc_bds_nodeb0x80cb-DFC_bds_NoDeb0x80cb.st ---- *)
(* --- Interface --- *)
{attribute 'external_name' := 'cmp_rts_DFC_bds_NoDeb0x80cb'}
TYPE DFC_bds_NoDeb0x80cb : STRUCT
		DTC            : UDINT := 16#80CB00;
		DFCid          : UINT  := 5;
		debounceMethod : USINT := TIME_IN_ROW;
	END_STRUCT
END_TYPE

(* ---- dfc_bds_nodeb0x80cc-DFC_bds_NoDeb0x80cc.st ---- *)
(* --- Interface --- *)
{attribute 'external_name' := 'cmp_rts_DFC_bds_NoDeb0x80cc'}
TYPE DFC_bds_NoDeb0x80cc : STRUCT
		DTC            : UDINT := 16#80CC00;
		DFCid          : UINT  := 6;
		debounceMethod : USINT := TIME_IN_ROW;
	END_STRUCT
END_TYPE

(* ---- dfc_bds_nodeb0x80cd-DFC_bds_NoDeb0x80cd.st ---- *)
(* --- Interface --- *)
{attribute 'external_name' := 'cmp_rts_DFC_bds_NoDeb0x80cd'}
TYPE DFC_bds_NoDeb0x80cd : STRUCT
		DTC            : UDINT := 16#80CD00;
		DFCid          : UINT  := 7;
		debounceMethod : USINT := TIME_IN_ROW;
	END_STRUCT
END_TYPE

(* ---- dfc_bds_nodeb0x80ce-DFC_bds_NoDeb0x80ce.st ---- *)
(* --- Interface --- *)
{attribute 'external_name' := 'cmp_rts_DFC_bds_NoDeb0x80ce'}
TYPE DFC_bds_NoDeb0x80ce : STRUCT
		DTC            : UDINT := 16#80CE00;
		DFCid          : UINT  := 8;
		debounceMethod : USINT := TIME_IN_ROW;
	END_STRUCT
END_TYPE

(* ---- dfc_bds_nodeb0x80cf-DFC_bds_NoDeb0x80cf.st ---- *)
(* --- Interface --- *)
{attribute 'external_name' := 'cmp_rts_DFC_bds_NoDeb0x80cf'}
TYPE DFC_bds_NoDeb0x80cf : STRUCT
		DTC            : UDINT := 16#80CF00;
		DFCid          : UINT  := 9;
		debounceMethod : USINT := TIME_IN_ROW;
	END_STRUCT
END_TYPE

(* ---- dfc_bds_nodeb0x80d0-DFC_bds_NoDeb0x80d0.st ---- *)
(* --- Interface --- *)
{attribute 'external_name' := 'cmp_rts_DFC_bds_NoDeb0x80d0'}
TYPE DFC_bds_NoDeb0x80d0 : STRUCT
		DTC            : UDINT := 16#80D000;
		DFCid          : UINT  := 10;
		debounceMethod : USINT := TIME_IN_ROW;
	END_STRUCT
END_TYPE

(* ---- dfc_bds_nodeb0x80d1-DFC_bds_NoDeb0x80d1.st ---- *)
(* --- Interface --- *)
{attribute 'external_name' := 'cmp_rts_DFC_bds_NoDeb0x80d1'}
TYPE DFC_bds_NoDeb0x80d1 : STRUCT
		DTC            : UDINT := 16#80D100;
		DFCid          : UINT  := 11;
		debounceMethod : USINT := TIME_IN_ROW;
	END_STRUCT
END_TYPE

(* ---- dfc_bds_nodeb0x80d2-DFC_bds_NoDeb0x80d2.st ---- *)
(* --- Interface --- *)
{attribute 'external_name' := 'cmp_rts_DFC_bds_NoDeb0x80d2'}
TYPE DFC_bds_NoDeb0x80d2 : STRUCT
		DTC            : UDINT := 16#80D200;
		DFCid          : UINT  := 12;
		debounceMethod : USINT := TIME_IN_ROW;
	END_STRUCT
END_TYPE

(* ---- dfc_bds_nodeb0x80d3-DFC_bds_NoDeb0x80d3.st ---- *)
(* --- Interface --- *)
{attribute 'external_name' := 'cmp_rts_DFC_bds_NoDeb0x80d3'}
TYPE DFC_bds_NoDeb0x80d3 : STRUCT
		DTC            : UDINT := 16#80D300;
		DFCid          : UINT  := 13;
		debounceMethod : USINT := TIME_IN_ROW;
	END_STRUCT
END_TYPE

(* ---- dfc_bds_nodeb0x80d4-DFC_bds_NoDeb0x80d4.st ---- *)
(* --- Interface --- *)
{attribute 'external_name' := 'cmp_rts_DFC_bds_NoDeb0x80d4'}
TYPE DFC_bds_NoDeb0x80d4 : STRUCT
		DTC            : UDINT := 16#80D400;
		DFCid          : UINT  := 14;
		debounceMethod : USINT := TIME_IN_ROW;
	END_STRUCT
END_TYPE

(* ---- dfc_bds_nodeb0x80d5-DFC_bds_NoDeb0x80d5.st ---- *)
(* --- Interface --- *)
{attribute 'external_name' := 'cmp_rts_DFC_bds_NoDeb0x80d5'}
TYPE DFC_bds_NoDeb0x80d5 : STRUCT
		DTC            : UDINT := 16#80D500;
		DFCid          : UINT  := 15;
		debounceMethod : USINT := TIME_IN_ROW;
	END_STRUCT
END_TYPE

(* ---- dfc_bds_nodeb0x80d6-DFC_bds_NoDeb0x80d6.st ---- *)
(* --- Interface --- *)
{attribute 'external_name' := 'cmp_rts_DFC_bds_NoDeb0x80d6'}
TYPE DFC_bds_NoDeb0x80d6 : STRUCT
		DTC            : UDINT := 16#80D600;
		DFCid          : UINT  := 16;
		debounceMethod : USINT := TIME_IN_ROW;
	END_STRUCT
END_TYPE

(* ---- dfc_bds_nodeb0x80d7-DFC_bds_NoDeb0x80d7.st ---- *)
(* --- Interface --- *)
{attribute 'external_name' := 'cmp_rts_DFC_bds_NoDeb0x80d7'}
TYPE DFC_bds_NoDeb0x80d7 : STRUCT
		DTC            : UDINT := 16#80D700;
		DFCid          : UINT  := 17;
		debounceMethod : USINT := TIME_IN_ROW;
	END_STRUCT
END_TYPE

(* ---- dfc_bds_nodeb0x80d8-DFC_bds_NoDeb0x80d8.st ---- *)
(* --- Interface --- *)
{attribute 'external_name' := 'cmp_rts_DFC_bds_NoDeb0x80d8'}
TYPE DFC_bds_NoDeb0x80d8 : STRUCT
		DTC            : UDINT := 16#80D800;
		DFCid          : UINT  := 18;
		debounceMethod : USINT := TIME_IN_ROW;
	END_STRUCT
END_TYPE

(* ---- dfc_bds_nodeb0x80d9-DFC_bds_NoDeb0x80d9.st ---- *)
(* --- Interface --- *)
{attribute 'external_name' := 'cmp_rts_DFC_bds_NoDeb0x80d9'}
TYPE DFC_bds_NoDeb0x80d9 : STRUCT
		DTC            : UDINT := 16#80D900;
		DFCid          : UINT  := 19;
		debounceMethod : USINT := TIME_IN_ROW;
	END_STRUCT
END_TYPE

(* ---- dfc_bds_nodeb0x80da-DFC_bds_NoDeb0x80da.st ---- *)
(* --- Interface --- *)
{attribute 'external_name' := 'cmp_rts_DFC_bds_NoDeb0x80da'}
TYPE DFC_bds_NoDeb0x80da : STRUCT
		DTC            : UDINT := 16#80DA00;
		DFCid          : UINT  := 20;
		debounceMethod : USINT := TIME_IN_ROW;
	END_STRUCT
END_TYPE

(* ---- dfc_bds_nodeb0x80db-DFC_bds_NoDeb0x80db.st ---- *)
(* --- Interface --- *)
{attribute 'external_name' := 'cmp_rts_DFC_bds_NoDeb0x80db'}
TYPE DFC_bds_NoDeb0x80db : STRUCT
		DTC            : UDINT := 16#80DB00;
		DFCid          : UINT  := 21;
		debounceMethod : USINT := TIME_IN_ROW;
	END_STRUCT
END_TYPE

(* ---- dfc_bds_nodeb0x80dc-DFC_bds_NoDeb0x80dc.st ---- *)
(* --- Interface --- *)
{attribute 'external_name' := 'cmp_rts_DFC_bds_NoDeb0x80dc'}
TYPE DFC_bds_NoDeb0x80dc : STRUCT
		DTC            : UDINT := 16#80DC00;
		DFCid          : UINT  := 22;
		debounceMethod : USINT := TIME_IN_ROW;
	END_STRUCT
END_TYPE

(* ---- dfc_bds_nodeb0x80dd-DFC_bds_NoDeb0x80dd.st ---- *)
(* --- Interface --- *)
{attribute 'external_name' := 'cmp_rts_DFC_bds_NoDeb0x80dd'}
TYPE DFC_bds_NoDeb0x80dd : STRUCT
		DTC            : UDINT := 16#80DD00;
		DFCid          : UINT  := 23;
		debounceMethod : USINT := TIME_IN_ROW;
	END_STRUCT
END_TYPE

(* ---- dfc_bds_nodeb0x80de-DFC_bds_NoDeb0x80de.st ---- *)
(* --- Interface --- *)
{attribute 'external_name' := 'cmp_rts_DFC_bds_NoDeb0x80de'}
TYPE DFC_bds_NoDeb0x80de : STRUCT
		DTC            : UDINT := 16#80DE00;
		DFCid          : UINT  := 24;
		debounceMethod : USINT := TIME_IN_ROW;
	END_STRUCT
END_TYPE

(* ---- dfc_bds_nodeb0x80df-DFC_bds_NoDeb0x80df.st ---- *)
(* --- Interface --- *)
{attribute 'external_name' := 'cmp_rts_DFC_bds_NoDeb0x80df'}
TYPE DFC_bds_NoDeb0x80df : STRUCT
		DTC            : UDINT := 16#80DF00;
		DFCid          : UINT  := 25;
		debounceMethod : USINT := TIME_IN_ROW;
	END_STRUCT
END_TYPE

(* ---- dfc_bds_nodeb0x80e0-DFC_bds_NoDeb0x80e0.st ---- *)
(* --- Interface --- *)
{attribute 'external_name' := 'cmp_rts_DFC_bds_NoDeb0x80e0'}
TYPE DFC_bds_NoDeb0x80e0 : STRUCT
		DTC            : UDINT := 16#80E000;
		DFCid          : UINT  := 26;
		debounceMethod : USINT := TIME_IN_ROW;
	END_STRUCT
END_TYPE

(* ---- dfc_bds_nodeb0x80e1-DFC_bds_NoDeb0x80e1.st ---- *)
(* --- Interface --- *)
{attribute 'external_name' := 'cmp_rts_DFC_bds_NoDeb0x80e1'}
TYPE DFC_bds_NoDeb0x80e1 : STRUCT
		DTC            : UDINT := 16#80E100;
		DFCid          : UINT  := 27;
		debounceMethod : USINT := TIME_IN_ROW;
	END_STRUCT
END_TYPE

(* ---- dfc_bds_nodeb0x80e2-DFC_bds_NoDeb0x80e2.st ---- *)
(* --- Interface --- *)
{attribute 'external_name' := 'cmp_rts_DFC_bds_NoDeb0x80e2'}
TYPE DFC_bds_NoDeb0x80e2 : STRUCT
		DTC            : UDINT := 16#80E200;
		DFCid          : UINT  := 28;
		debounceMethod : USINT := TIME_IN_ROW;
	END_STRUCT
END_TYPE

(* ---- dfc_bds_nodeb0x80e3-DFC_bds_NoDeb0x80e3.st ---- *)
(* --- Interface --- *)
{attribute 'external_name' := 'cmp_rts_DFC_bds_NoDeb0x80e3'}
TYPE DFC_bds_NoDeb0x80e3 : STRUCT
		DTC            : UDINT := 16#80E300;
		DFCid          : UINT  := 29;
		debounceMethod : USINT := TIME_IN_ROW;
	END_STRUCT
END_TYPE

(* ---- dfc_bds_nodeb0x80e4-DFC_bds_NoDeb0x80e4.st ---- *)
(* --- Interface --- *)
{attribute 'external_name' := 'cmp_rts_DFC_bds_NoDeb0x80e4'}
TYPE DFC_bds_NoDeb0x80e4 : STRUCT
		DTC            : UDINT := 16#80E400;
		DFCid          : UINT  := 30;
		debounceMethod : USINT := TIME_IN_ROW;
	END_STRUCT
END_TYPE

(* ---- dfc_bds_nodeb0x80e5-DFC_bds_NoDeb0x80e5.st ---- *)
(* --- Interface --- *)
{attribute 'external_name' := 'cmp_rts_DFC_bds_NoDeb0x80e5'}
TYPE DFC_bds_NoDeb0x80e5 : STRUCT
		DTC            : UDINT := 16#80E500;
		DFCid          : UINT  := 31;
		debounceMethod : USINT := TIME_IN_ROW;
	END_STRUCT
END_TYPE

(* ---- dfc_bds_nodeb0x80e6-DFC_bds_NoDeb0x80e6.st ---- *)
(* --- Interface --- *)
{attribute 'external_name' := 'cmp_rts_DFC_bds_NoDeb0x80e6'}
TYPE DFC_bds_NoDeb0x80e6 : STRUCT
		DTC            : UDINT := 16#80E600;
		DFCid          : UINT  := 32;
		debounceMethod : USINT := TIME_IN_ROW;
	END_STRUCT
END_TYPE

(* ---- dfc_bds_nodeb0x80e7-DFC_bds_NoDeb0x80e7.st ---- *)
(* --- Interface --- *)
{attribute 'external_name' := 'cmp_rts_DFC_bds_NoDeb0x80e7'}
TYPE DFC_bds_NoDeb0x80e7 : STRUCT
		DTC            : UDINT := 16#80E700;
		DFCid          : UINT  := 33;
		debounceMethod : USINT := TIME_IN_ROW;
	END_STRUCT
END_TYPE

(* ---- dfc_bds_nodeb0x80e8-DFC_bds_NoDeb0x80e8.st ---- *)
(* --- Interface --- *)
{attribute 'external_name' := 'cmp_rts_DFC_bds_NoDeb0x80e8'}
TYPE DFC_bds_NoDeb0x80e8 : STRUCT
		DTC            : UDINT := 16#80E800;
		DFCid          : UINT  := 34;
		debounceMethod : USINT := TIME_IN_ROW;
	END_STRUCT
END_TYPE

(* ---- dfc_bds_nodeb0x80e9-DFC_bds_NoDeb0x80e9.st ---- *)
(* --- Interface --- *)
{attribute 'external_name' := 'cmp_rts_DFC_bds_NoDeb0x80e9'}
TYPE DFC_bds_NoDeb0x80e9 : STRUCT
		DTC            : UDINT := 16#80E900;
		DFCid          : UINT  := 35;
		debounceMethod : USINT := TIME_IN_ROW;
	END_STRUCT
END_TYPE

(* ---- dfc_bds_nodeb0x80ea-DFC_bds_NoDeb0x80ea.st ---- *)
(* --- Interface --- *)
{attribute 'external_name' := 'cmp_rts_DFC_bds_NoDeb0x80ea'}
TYPE DFC_bds_NoDeb0x80ea : STRUCT
		DTC            : UDINT := 16#80EA00;
		DFCid          : UINT  := 36;
		debounceMethod : USINT := TIME_IN_ROW;
	END_STRUCT
END_TYPE

(* ---- dfc_bds_nodeb0x80eb-DFC_bds_NoDeb0x80eb.st ---- *)
(* --- Interface --- *)
{attribute 'external_name' := 'cmp_rts_DFC_bds_NoDeb0x80eb'}
TYPE DFC_bds_NoDeb0x80eb : STRUCT
		DTC            : UDINT := 16#80EB00;
		DFCid          : UINT  := 37;
		debounceMethod : USINT := TIME_IN_ROW;
	END_STRUCT
END_TYPE

(* ---- dfc_bds_nodeb0x80ec-DFC_bds_NoDeb0x80ec.st ---- *)
(* --- Interface --- *)
{attribute 'external_name' := 'cmp_rts_DFC_bds_NoDeb0x80ec'}
TYPE DFC_bds_NoDeb0x80ec : STRUCT
		DTC            : UDINT := 16#80EC00;
		DFCid          : UINT  := 38;
		debounceMethod : USINT := TIME_IN_ROW;
	END_STRUCT
END_TYPE

(* ---- dfc_bds_nodeb0x80ed-DFC_bds_NoDeb0x80ed.st ---- *)
(* --- Interface --- *)
{attribute 'external_name' := 'cmp_rts_DFC_bds_NoDeb0x80ed'}
TYPE DFC_bds_NoDeb0x80ed : STRUCT
		DTC            : UDINT := 16#80ED00;
		DFCid          : UINT  := 39;
		debounceMethod : USINT := TIME_IN_ROW;
	END_STRUCT
END_TYPE

(* ---- dfc_bds_nodeb0x80ee-DFC_bds_NoDeb0x80ee.st ---- *)
(* --- Interface --- *)
{attribute 'external_name' := 'cmp_rts_DFC_bds_NoDeb0x80ee'}
TYPE DFC_bds_NoDeb0x80ee : STRUCT
		DTC            : UDINT := 16#80EE00;
		DFCid          : UINT  := 40;
		debounceMethod : USINT := TIME_IN_ROW;
	END_STRUCT
END_TYPE

(* ---- dfc_bds_nodeb0x80ef-DFC_bds_NoDeb0x80ef.st ---- *)
(* --- Interface --- *)
{attribute 'external_name' := 'cmp_rts_DFC_bds_NoDeb0x80ef'}
TYPE DFC_bds_NoDeb0x80ef : STRUCT
		DTC            : UDINT := 16#80EF00;
		DFCid          : UINT  := 41;
		debounceMethod : USINT := TIME_IN_ROW;
	END_STRUCT
END_TYPE

(* ---- dfc_bds_nodeb0x80f0-DFC_bds_NoDeb0x80f0.st ---- *)
(* --- Interface --- *)
{attribute 'external_name' := 'cmp_rts_DFC_bds_NoDeb0x80f0'}
TYPE DFC_bds_NoDeb0x80f0 : STRUCT
		DTC            : UDINT := 16#80F000;
		DFCid          : UINT  := 42;
		debounceMethod : USINT := TIME_IN_ROW;
	END_STRUCT
END_TYPE

(* ---- dfc_bds_nodeb0x80f1-DFC_bds_NoDeb0x80f1.st ---- *)
(* --- Interface --- *)
{attribute 'external_name' := 'cmp_rts_DFC_bds_NoDeb0x80f1'}
TYPE DFC_bds_NoDeb0x80f1 : STRUCT
		DTC            : UDINT := 16#80F100;
		DFCid          : UINT  := 43;
		debounceMethod : USINT := TIME_IN_ROW;
	END_STRUCT
END_TYPE

(* ---- dfc_bds_nodeb0x80f2-DFC_bds_NoDeb0x80f2.st ---- *)
(* --- Interface --- *)
{attribute 'external_name' := 'cmp_rts_DFC_bds_NoDeb0x80f2'}
TYPE DFC_bds_NoDeb0x80f2 : STRUCT
		DTC            : UDINT := 16#80F200;
		DFCid          : UINT  := 44;
		debounceMethod : USINT := TIME_IN_ROW;
	END_STRUCT
END_TYPE

(* ---- dfc_bds_nodeb0x80f3-DFC_bds_NoDeb0x80f3.st ---- *)
(* --- Interface --- *)
{attribute 'external_name' := 'cmp_rts_DFC_bds_NoDeb0x80f3'}
TYPE DFC_bds_NoDeb0x80f3 : STRUCT
		DTC            : UDINT := 16#80F300;
		DFCid          : UINT  := 45;
		debounceMethod : USINT := TIME_IN_ROW;
	END_STRUCT
END_TYPE

(* ---- dfc_bds_nodeb0x80f4-DFC_bds_NoDeb0x80f4.st ---- *)
(* --- Interface --- *)
{attribute 'external_name' := 'cmp_rts_DFC_bds_NoDeb0x80f4'}
TYPE DFC_bds_NoDeb0x80f4 : STRUCT
		DTC            : UDINT := 16#80F400;
		DFCid          : UINT  := 46;
		debounceMethod : USINT := TIME_IN_ROW;
	END_STRUCT
END_TYPE

(* ---- dfc_bds_nodeb0x80f5-DFC_bds_NoDeb0x80f5.st ---- *)
(* --- Interface --- *)
{attribute 'external_name' := 'cmp_rts_DFC_bds_NoDeb0x80f5'}
TYPE DFC_bds_NoDeb0x80f5 : STRUCT
		DTC            : UDINT := 16#80F500;
		DFCid          : UINT  := 47;
		debounceMethod : USINT := TIME_IN_ROW;
	END_STRUCT
END_TYPE

(* ---- dfc_bds_nodeb0x80f6-DFC_bds_NoDeb0x80f6.st ---- *)
(* --- Interface --- *)
{attribute 'external_name' := 'cmp_rts_DFC_bds_NoDeb0x80f6'}
TYPE DFC_bds_NoDeb0x80f6 : STRUCT
		DTC            : UDINT := 16#80F600;
		DFCid          : UINT  := 48;
		debounceMethod : USINT := TIME_IN_ROW;
	END_STRUCT
END_TYPE

(* ---- dfc_bds_nodeb0x80f7-DFC_bds_NoDeb0x80f7.st ---- *)
(* --- Interface --- *)
{attribute 'external_name' := 'cmp_rts_DFC_bds_NoDeb0x80f7'}
TYPE DFC_bds_NoDeb0x80f7 : STRUCT
		DTC            : UDINT := 16#80F700;
		DFCid          : UINT  := 49;
		debounceMethod : USINT := TIME_IN_ROW;
	END_STRUCT
END_TYPE

(* ---- dfc_bds_nodeb0x80f8-DFC_bds_NoDeb0x80f8.st ---- *)
(* --- Interface --- *)
{attribute 'external_name' := 'cmp_rts_DFC_bds_NoDeb0x80f8'}
TYPE DFC_bds_NoDeb0x80f8 : STRUCT
		DTC            : UDINT := 16#80F800;
		DFCid          : UINT  := 50;
		debounceMethod : USINT := TIME_IN_ROW;
	END_STRUCT
END_TYPE

(* ---- dfc_bds_nodeb0x80f9-DFC_bds_NoDeb0x80f9.st ---- *)
(* --- Interface --- *)
{attribute 'external_name' := 'cmp_rts_DFC_bds_NoDeb0x80f9'}
TYPE DFC_bds_NoDeb0x80f9 : STRUCT
		DTC            : UDINT := 16#80F900;
		DFCid          : UINT  := 51;
		debounceMethod : USINT := TIME_IN_ROW;
	END_STRUCT
END_TYPE

(* ---- dfc_bds_nodeb0x80fa-DFC_bds_NoDeb0x80fa.st ---- *)
(* --- Interface --- *)
{attribute 'external_name' := 'cmp_rts_DFC_bds_NoDeb0x80fa'}
TYPE DFC_bds_NoDeb0x80fa : STRUCT
		DTC            : UDINT := 16#80FA00;
		DFCid          : UINT  := 52;
		debounceMethod : USINT := TIME_IN_ROW;
	END_STRUCT
END_TYPE

(* ---- dfc_bds_nodeb0x80fb-DFC_bds_NoDeb0x80fb.st ---- *)
(* --- Interface --- *)
{attribute 'external_name' := 'cmp_rts_DFC_bds_NoDeb0x80fb'}
TYPE DFC_bds_NoDeb0x80fb : STRUCT
		DTC            : UDINT := 16#80FB00;
		DFCid          : UINT  := 53;
		debounceMethod : USINT := TIME_IN_ROW;
	END_STRUCT
END_TYPE

(* ---- dfc_bds_nodeb0x80fc-DFC_bds_NoDeb0x80fc.st ---- *)
(* --- Interface --- *)
{attribute 'external_name' := 'cmp_rts_DFC_bds_NoDeb0x80fc'}
TYPE DFC_bds_NoDeb0x80fc : STRUCT
		DTC            : UDINT := 16#80FC00;
		DFCid          : UINT  := 54;
		debounceMethod : USINT := TIME_IN_ROW;
	END_STRUCT
END_TYPE

(* ---- dfc_bds_nodeb0x80fd-DFC_bds_NoDeb0x80fd.st ---- *)
(* --- Interface --- *)
{attribute 'external_name' := 'cmp_rts_DFC_bds_NoDeb0x80fd'}
TYPE DFC_bds_NoDeb0x80fd : STRUCT
		DTC            : UDINT := 16#80FD00;
		DFCid          : UINT  := 55;
		debounceMethod : USINT := TIME_IN_ROW;
	END_STRUCT
END_TYPE

(* ---- dfc_bds_nodeb0x80fe-DFC_bds_NoDeb0x80fe.st ---- *)
(* --- Interface --- *)
{attribute 'external_name' := 'cmp_rts_DFC_bds_NoDeb0x80fe'}
TYPE DFC_bds_NoDeb0x80fe : STRUCT
		DTC            : UDINT := 16#80FE00;
		DFCid          : UINT  := 56;
		debounceMethod : USINT := TIME_IN_ROW;
	END_STRUCT
END_TYPE

(* ---- dfc_bds_nodeb0x80ff-DFC_bds_NoDeb0x80ff.st ---- *)
(* --- Interface --- *)
{attribute 'external_name' := 'cmp_rts_DFC_bds_NoDeb0x80ff'}
TYPE DFC_bds_NoDeb0x80ff : STRUCT
		DTC            : UDINT := 16#80FF00;
		DFCid          : UINT  := 57;
		debounceMethod : USINT := TIME_IN_ROW;
	END_STRUCT
END_TYPE

(* ---- dfc_bds_nodeb0x8100-DFC_bds_NoDeb0x8100.st ---- *)
(* --- Interface --- *)
{attribute 'external_name' := 'cmp_rts_DFC_bds_NoDeb0x8100'}
TYPE DFC_bds_NoDeb0x8100 : STRUCT
		DTC            : UDINT := 16#810000;
		DFCid          : UINT  := 58;
		debounceMethod : USINT := TIME_IN_ROW;
	END_STRUCT
END_TYPE

(* ---- dfc_bds_nodeb0x8101-DFC_bds_NoDeb0x8101.st ---- *)
(* --- Interface --- *)
{attribute 'external_name' := 'cmp_rts_DFC_bds_NoDeb0x8101'}
TYPE DFC_bds_NoDeb0x8101 : STRUCT
		DTC            : UDINT := 16#810100;
		DFCid          : UINT  := 59;
		debounceMethod : USINT := TIME_IN_ROW;
	END_STRUCT
END_TYPE

(* ---- dfc_bds_nodeb0x8102-DFC_bds_NoDeb0x8102.st ---- *)
(* --- Interface --- *)
{attribute 'external_name' := 'cmp_rts_DFC_bds_NoDeb0x8102'}
TYPE DFC_bds_NoDeb0x8102 : STRUCT
		DTC            : UDINT := 16#810200;
		DFCid          : UINT  := 60;
		debounceMethod : USINT := TIME_IN_ROW;
	END_STRUCT
END_TYPE

(* ---- dfc_bds_nodeb0x8103-DFC_bds_NoDeb0x8103.st ---- *)
(* --- Interface --- *)
{attribute 'external_name' := 'cmp_rts_DFC_bds_NoDeb0x8103'}
TYPE DFC_bds_NoDeb0x8103 : STRUCT
		DTC            : UDINT := 16#810300;
		DFCid          : UINT  := 61;
		debounceMethod : USINT := TIME_IN_ROW;
	END_STRUCT
END_TYPE

(* ---- dfc_bds_nodeb0x8104-DFC_bds_NoDeb0x8104.st ---- *)
(* --- Interface --- *)
{attribute 'external_name' := 'cmp_rts_DFC_bds_NoDeb0x8104'}
TYPE DFC_bds_NoDeb0x8104 : STRUCT
		DTC            : UDINT := 16#810400;
		DFCid          : UINT  := 62;
		debounceMethod : USINT := TIME_IN_ROW;
	END_STRUCT
END_TYPE

(* ---- dfc_bds_nodeb0x8105-DFC_bds_NoDeb0x8105.st ---- *)
(* --- Interface --- *)
{attribute 'external_name' := 'cmp_rts_DFC_bds_NoDeb0x8105'}
TYPE DFC_bds_NoDeb0x8105 : STRUCT
		DTC            : UDINT := 16#810500;
		DFCid          : UINT  := 63;
		debounceMethod : USINT := TIME_IN_ROW;
	END_STRUCT
END_TYPE

(* ---- dfc_bds_nodeb0x8106-DFC_bds_NoDeb0x8106.st ---- *)
(* --- Interface --- *)
{attribute 'external_name' := 'cmp_rts_DFC_bds_NoDeb0x8106'}
TYPE DFC_bds_NoDeb0x8106 : STRUCT
		DTC            : UDINT := 16#810600;
		DFCid          : UINT  := 64;
		debounceMethod : USINT := TIME_IN_ROW;
	END_STRUCT
END_TYPE

(* ---- dfc_bds_nodeb0x8107-DFC_bds_NoDeb0x8107.st ---- *)
(* --- Interface --- *)
{attribute 'external_name' := 'cmp_rts_DFC_bds_NoDeb0x8107'}
TYPE DFC_bds_NoDeb0x8107 : STRUCT
		DTC            : UDINT := 16#810700;
		DFCid          : UINT  := 65;
		debounceMethod : USINT := TIME_IN_ROW;
	END_STRUCT
END_TYPE

(* ---- dfc_bds_nodeb0x8108-DFC_bds_NoDeb0x8108.st ---- *)
(* --- Interface --- *)
{attribute 'external_name' := 'cmp_rts_DFC_bds_NoDeb0x8108'}
TYPE DFC_bds_NoDeb0x8108 : STRUCT
		DTC            : UDINT := 16#810800;
		DFCid          : UINT  := 66;
		debounceMethod : USINT := TIME_IN_ROW;
	END_STRUCT
END_TYPE

(* ---- dfc_bds_nodeb0x8109-DFC_bds_NoDeb0x8109.st ---- *)
(* --- Interface --- *)
{attribute 'external_name' := 'cmp_rts_DFC_bds_NoDeb0x8109'}
TYPE DFC_bds_NoDeb0x8109 : STRUCT
		DTC            : UDINT := 16#810900;
		DFCid          : UINT  := 67;
		debounceMethod : USINT := TIME_IN_ROW;
	END_STRUCT
END_TYPE

(* ---- dfc_bds_nodeb0x810a-DFC_bds_NoDeb0x810a.st ---- *)
(* --- Interface --- *)
{attribute 'external_name' := 'cmp_rts_DFC_bds_NoDeb0x810a'}
TYPE DFC_bds_NoDeb0x810a : STRUCT
		DTC            : UDINT := 16#810A00;
		DFCid          : UINT  := 68;
		debounceMethod : USINT := TIME_IN_ROW;
	END_STRUCT
END_TYPE

(* ---- dfc_bds_nodeb0x810b-DFC_bds_NoDeb0x810b.st ---- *)
(* --- Interface --- *)
{attribute 'external_name' := 'cmp_rts_DFC_bds_NoDeb0x810b'}
TYPE DFC_bds_NoDeb0x810b : STRUCT
		DTC            : UDINT := 16#810B00;
		DFCid          : UINT  := 69;
		debounceMethod : USINT := TIME_IN_ROW;
	END_STRUCT
END_TYPE

(* ---- dfc_bds_nodeb0x810c-DFC_bds_NoDeb0x810c.st ---- *)
(* --- Interface --- *)
{attribute 'external_name' := 'cmp_rts_DFC_bds_NoDeb0x810c'}
TYPE DFC_bds_NoDeb0x810c : STRUCT
		DTC            : UDINT := 16#810C00;
		DFCid          : UINT  := 70;
		debounceMethod : USINT := TIME_IN_ROW;
	END_STRUCT
END_TYPE

(* ---- dfc_bds_nodeb0x810d-DFC_bds_NoDeb0x810d.st ---- *)
(* --- Interface --- *)
{attribute 'external_name' := 'cmp_rts_DFC_bds_NoDeb0x810d'}
TYPE DFC_bds_NoDeb0x810d : STRUCT
		DTC            : UDINT := 16#810D00;
		DFCid          : UINT  := 71;
		debounceMethod : USINT := TIME_IN_ROW;
	END_STRUCT
END_TYPE

(* ---- dfc_bds_nodeb0x810e-DFC_bds_NoDeb0x810e.st ---- *)
(* --- Interface --- *)
{attribute 'external_name' := 'cmp_rts_DFC_bds_NoDeb0x810e'}
TYPE DFC_bds_NoDeb0x810e : STRUCT
		DTC            : UDINT := 16#810E00;
		DFCid          : UINT  := 72;
		debounceMethod : USINT := TIME_IN_ROW;
	END_STRUCT
END_TYPE

(* ---- dfc_bds_nodeb0x810f-DFC_bds_NoDeb0x810f.st ---- *)
(* --- Interface --- *)
{attribute 'external_name' := 'cmp_rts_DFC_bds_NoDeb0x810f'}
TYPE DFC_bds_NoDeb0x810f : STRUCT
		DTC            : UDINT := 16#810F00;
		DFCid          : UINT  := 73;
		debounceMethod : USINT := TIME_IN_ROW;
	END_STRUCT
END_TYPE

(* ---- dfc_bds_nodeb0x8110-DFC_bds_NoDeb0x8110.st ---- *)
(* --- Interface --- *)
{attribute 'external_name' := 'cmp_rts_DFC_bds_NoDeb0x8110'}
TYPE DFC_bds_NoDeb0x8110 : STRUCT
		DTC            : UDINT := 16#811000;
		DFCid          : UINT  := 74;
		debounceMethod : USINT := TIME_IN_ROW;
	END_STRUCT
END_TYPE

(* ---- dfc_bds_nodeb0x8111-DFC_bds_NoDeb0x8111.st ---- *)
(* --- Interface --- *)
{attribute 'external_name' := 'cmp_rts_DFC_bds_NoDeb0x8111'}
TYPE DFC_bds_NoDeb0x8111 : STRUCT
		DTC            : UDINT := 16#811100;
		DFCid          : UINT  := 75;
		debounceMethod : USINT := TIME_IN_ROW;
	END_STRUCT
END_TYPE

(* ---- dfc_bds_nodeb0x8112-DFC_bds_NoDeb0x8112.st ---- *)
(* --- Interface --- *)
{attribute 'external_name' := 'cmp_rts_DFC_bds_NoDeb0x8112'}
TYPE DFC_bds_NoDeb0x8112 : STRUCT
		DTC            : UDINT := 16#811200;
		DFCid          : UINT  := 76;
		debounceMethod : USINT := TIME_IN_ROW;
	END_STRUCT
END_TYPE

(* ---- dfc_bds_nodeb0x8113-DFC_bds_NoDeb0x8113.st ---- *)
(* --- Interface --- *)
{attribute 'external_name' := 'cmp_rts_DFC_bds_NoDeb0x8113'}
TYPE DFC_bds_NoDeb0x8113 : STRUCT
		DTC            : UDINT := 16#811300;
		DFCid          : UINT  := 77;
		debounceMethod : USINT := TIME_IN_ROW;
	END_STRUCT
END_TYPE

(* ---- dfc_bds_nodeb0x8114-DFC_bds_NoDeb0x8114.st ---- *)
(* --- Interface --- *)
{attribute 'external_name' := 'cmp_rts_DFC_bds_NoDeb0x8114'}
TYPE DFC_bds_NoDeb0x8114 : STRUCT
		DTC            : UDINT := 16#811400;
		DFCid          : UINT  := 78;
		debounceMethod : USINT := TIME_IN_ROW;
	END_STRUCT
END_TYPE

(* ---- dfc_bds_nodeb0x8115-DFC_bds_NoDeb0x8115.st ---- *)
(* --- Interface --- *)
{attribute 'external_name' := 'cmp_rts_DFC_bds_NoDeb0x8115'}
TYPE DFC_bds_NoDeb0x8115 : STRUCT
		DTC            : UDINT := 16#811500;
		DFCid          : UINT  := 79;
		debounceMethod : USINT := TIME_IN_ROW;
	END_STRUCT
END_TYPE

(* ---- dfc_bds_nodeb0x8116-DFC_bds_NoDeb0x8116.st ---- *)
(* --- Interface --- *)
{attribute 'external_name' := 'cmp_rts_DFC_bds_NoDeb0x8116'}
TYPE DFC_bds_NoDeb0x8116 : STRUCT
		DTC            : UDINT := 16#811600;
		DFCid          : UINT  := 80;
		debounceMethod : USINT := TIME_IN_ROW;
	END_STRUCT
END_TYPE

(* ---- dfc_bds_nodeb0x8117-DFC_bds_NoDeb0x8117.st ---- *)
(* --- Interface --- *)
{attribute 'external_name' := 'cmp_rts_DFC_bds_NoDeb0x8117'}
TYPE DFC_bds_NoDeb0x8117 : STRUCT
		DTC            : UDINT := 16#811700;
		DFCid          : UINT  := 81;
		debounceMethod : USINT := TIME_IN_ROW;
	END_STRUCT
END_TYPE

(* ---- dfc_bds_nodeb0x8118-DFC_bds_NoDeb0x8118.st ---- *)
(* --- Interface --- *)
{attribute 'external_name' := 'cmp_rts_DFC_bds_NoDeb0x8118'}
TYPE DFC_bds_NoDeb0x8118 : STRUCT
		DTC            : UDINT := 16#811800;
		DFCid          : UINT  := 82;
		debounceMethod : USINT := TIME_IN_ROW;
	END_STRUCT
END_TYPE

(* ---- dfc_bds_nodeb0x8119-DFC_bds_NoDeb0x8119.st ---- *)
(* --- Interface --- *)
{attribute 'external_name' := 'cmp_rts_DFC_bds_NoDeb0x8119'}
TYPE DFC_bds_NoDeb0x8119 : STRUCT
		DTC            : UDINT := 16#811900;
		DFCid          : UINT  := 83;
		debounceMethod : USINT := TIME_IN_ROW;
	END_STRUCT
END_TYPE

(* ---- dfc_bds_nodeb0x811a-DFC_bds_NoDeb0x811a.st ---- *)
(* --- Interface --- *)
{attribute 'external_name' := 'cmp_rts_DFC_bds_NoDeb0x811a'}
TYPE DFC_bds_NoDeb0x811a : STRUCT
		DTC            : UDINT := 16#811A00;
		DFCid          : UINT  := 84;
		debounceMethod : USINT := TIME_IN_ROW;
	END_STRUCT
END_TYPE

(* ---- dfc_bds_nodeb0x811b-DFC_bds_NoDeb0x811b.st ---- *)
(* --- Interface --- *)
{attribute 'external_name' := 'cmp_rts_DFC_bds_NoDeb0x811b'}
TYPE DFC_bds_NoDeb0x811b : STRUCT
		DTC            : UDINT := 16#811B00;
		DFCid          : UINT  := 85;
		debounceMethod : USINT := TIME_IN_ROW;
	END_STRUCT
END_TYPE

(* ---- dfc_bds_nodeb0x811c-DFC_bds_NoDeb0x811c.st ---- *)
(* --- Interface --- *)
{attribute 'external_name' := 'cmp_rts_DFC_bds_NoDeb0x811c'}
TYPE DFC_bds_NoDeb0x811c : STRUCT
		DTC            : UDINT := 16#811C00;
		DFCid          : UINT  := 86;
		debounceMethod : USINT := TIME_IN_ROW;
	END_STRUCT
END_TYPE

(* ---- dfc_bds_nodeb0x811d-DFC_bds_NoDeb0x811d.st ---- *)
(* --- Interface --- *)
{attribute 'external_name' := 'cmp_rts_DFC_bds_NoDeb0x811d'}
TYPE DFC_bds_NoDeb0x811d : STRUCT
		DTC            : UDINT := 16#811D00;
		DFCid          : UINT  := 87;
		debounceMethod : USINT := TIME_IN_ROW;
	END_STRUCT
END_TYPE

(* ---- dfc_bds_nodeb0x811e-DFC_bds_NoDeb0x811e.st ---- *)
(* --- Interface --- *)
{attribute 'external_name' := 'cmp_rts_DFC_bds_NoDeb0x811e'}
TYPE DFC_bds_NoDeb0x811e : STRUCT
		DTC            : UDINT := 16#811E00;
		DFCid          : UINT  := 88;
		debounceMethod : USINT := TIME_IN_ROW;
	END_STRUCT
END_TYPE

(* ---- dfc_bds_nodeb0x811f-DFC_bds_NoDeb0x811f.st ---- *)
(* --- Interface --- *)
{attribute 'external_name' := 'cmp_rts_DFC_bds_NoDeb0x811f'}
TYPE DFC_bds_NoDeb0x811f : STRUCT
		DTC            : UDINT := 16#811F00;
		DFCid          : UINT  := 89;
		debounceMethod : USINT := TIME_IN_ROW;
	END_STRUCT
END_TYPE

(* ---- dfc_bds_nodeb0x8120-DFC_bds_NoDeb0x8120.st ---- *)
(* --- Interface --- *)
{attribute 'external_name' := 'cmp_rts_DFC_bds_NoDeb0x8120'}
TYPE DFC_bds_NoDeb0x8120 : STRUCT
		DTC            : UDINT := 16#812000;
		DFCid          : UINT  := 90;
		debounceMethod : USINT := TIME_IN_ROW;
	END_STRUCT
END_TYPE

(* ---- dfc_bds_nodeb0x8121-DFC_bds_NoDeb0x8121.st ---- *)
(* --- Interface --- *)
{attribute 'external_name' := 'cmp_rts_DFC_bds_NoDeb0x8121'}
TYPE DFC_bds_NoDeb0x8121 : STRUCT
		DTC            : UDINT := 16#812100;
		DFCid          : UINT  := 91;
		debounceMethod : USINT := TIME_IN_ROW;
	END_STRUCT
END_TYPE

(* ---- dfc_bds_nodeb0x8122-DFC_bds_NoDeb0x8122.st ---- *)
(* --- Interface --- *)
{attribute 'external_name' := 'cmp_rts_DFC_bds_NoDeb0x8122'}
TYPE DFC_bds_NoDeb0x8122 : STRUCT
		DTC            : UDINT := 16#812200;
		DFCid          : UINT  := 92;
		debounceMethod : USINT := TIME_IN_ROW;
	END_STRUCT
END_TYPE

(* ---- dfc_bds_nodeb0x8123-DFC_bds_NoDeb0x8123.st ---- *)
(* --- Interface --- *)
{attribute 'external_name' := 'cmp_rts_DFC_bds_NoDeb0x8123'}
TYPE DFC_bds_NoDeb0x8123 : STRUCT
		DTC            : UDINT := 16#812300;
		DFCid          : UINT  := 93;
		debounceMethod : USINT := TIME_IN_ROW;
	END_STRUCT
END_TYPE

(* ---- dfc_bds_nodeb0x8124-DFC_bds_NoDeb0x8124.st ---- *)
(* --- Interface --- *)
{attribute 'external_name' := 'cmp_rts_DFC_bds_NoDeb0x8124'}
TYPE DFC_bds_NoDeb0x8124 : STRUCT
		DTC            : UDINT := 16#812400;
		DFCid          : UINT  := 94;
		debounceMethod : USINT := TIME_IN_ROW;
	END_STRUCT
END_TYPE

(* ---- dfc_bds_nodeb0x8125-DFC_bds_NoDeb0x8125.st ---- *)
(* --- Interface --- *)
{attribute 'external_name' := 'cmp_rts_DFC_bds_NoDeb0x8125'}
TYPE DFC_bds_NoDeb0x8125 : STRUCT
		DTC            : UDINT := 16#812500;
		DFCid          : UINT  := 95;
		debounceMethod : USINT := TIME_IN_ROW;
	END_STRUCT
END_TYPE

(* ---- dfc_bds_nodeb0x8126-DFC_bds_NoDeb0x8126.st ---- *)
(* --- Interface --- *)
{attribute 'external_name' := 'cmp_rts_DFC_bds_NoDeb0x8126'}
TYPE DFC_bds_NoDeb0x8126 : STRUCT
		DTC            : UDINT := 16#812600;
		DFCid          : UINT  := 96;
		debounceMethod : USINT := TIME_IN_ROW;
	END_STRUCT
END_TYPE

(* ---- dfc_bds_nodeb0x8127-DFC_bds_NoDeb0x8127.st ---- *)
(* --- Interface --- *)
{attribute 'external_name' := 'cmp_rts_DFC_bds_NoDeb0x8127'}
TYPE DFC_bds_NoDeb0x8127 : STRUCT
		DTC            : UDINT := 16#812700;
		DFCid          : UINT  := 97;
		debounceMethod : USINT := TIME_IN_ROW;
	END_STRUCT
END_TYPE

(* ---- dfc_bds_nodeb0x8128-DFC_bds_NoDeb0x8128.st ---- *)
(* --- Interface --- *)
{attribute 'external_name' := 'cmp_rts_DFC_bds_NoDeb0x8128'}
TYPE DFC_bds_NoDeb0x8128 : STRUCT
		DTC            : UDINT := 16#812800;
		DFCid          : UINT  := 98;
		debounceMethod : USINT := TIME_IN_ROW;
	END_STRUCT
END_TYPE

(* ---- dfc_bds_nodeb0x8129-DFC_bds_NoDeb0x8129.st ---- *)
(* --- Interface --- *)
{attribute 'external_name' := 'cmp_rts_DFC_bds_NoDeb0x8129'}
TYPE DFC_bds_NoDeb0x8129 : STRUCT
		DTC            : UDINT := 16#812900;
		DFCid          : UINT  := 99;
		debounceMethod : USINT := TIME_IN_ROW;
	END_STRUCT
END_TYPE

(* ---- dfc_bds_nodeb0x812a-DFC_bds_NoDeb0x812a.st ---- *)
(* --- Interface --- *)
{attribute 'external_name' := 'cmp_rts_DFC_bds_NoDeb0x812a'}
TYPE DFC_bds_NoDeb0x812a : STRUCT
		DTC            : UDINT := 16#812A00;
		DFCid          : UINT  := 100;
		debounceMethod : USINT := TIME_IN_ROW;
	END_STRUCT
END_TYPE

(* ---- dfc_bds_nodeb0x8c01-DFC_bds_NoDeb0x8C01.st ---- *)
(* --- Interface --- *)
{attribute 'external_name' := 'cmp_rts_DFC_bds_NoDeb0x8C01'}
TYPE DFC_bds_NoDeb0x8C01 : STRUCT
		DTC            : UDINT := 16#8C0100;
		DFCid          : UINT  := 820;
		debounceMethod : USINT := NO_DEBOUNCE;
	END_STRUCT
END_TYPE

(* ---- dfc_bds_nodeb0x8c02-DFC_bds_NoDeb0x8C02.st ---- *)
(* --- Interface --- *)
{attribute 'external_name' := 'cmp_rts_DFC_bds_NoDeb0x8C02'}
TYPE DFC_bds_NoDeb0x8C02 : STRUCT
		DTC            : UDINT := 16#8C0200;
		DFCid          : UINT  := 821;
		debounceMethod : USINT := NO_DEBOUNCE;
	END_STRUCT
END_TYPE

(* ---- dfc_bds_nodeb0x8c03-DFC_bds_NoDeb0x8C03.st ---- *)
(* --- Interface --- *)
{attribute 'external_name' := 'cmp_rts_DFC_bds_NoDeb0x8C03'}
TYPE DFC_bds_NoDeb0x8C03 : STRUCT
		DTC            : UDINT := 16#8C0300;
		DFCid          : UINT  := 822;
		debounceMethod : USINT := NO_DEBOUNCE;
	END_STRUCT
END_TYPE

(* ---- dfc_bds_tiinrow0x8b01-DFC_bds_TiInRow0x8B01.st ---- *)
(* --- Interface --- *)
{attribute 'external_name' := 'cmp_rts_DFC_bds_TiInRow0x8B01'}
TYPE DFC_bds_TiInRow0x8B01 : STRUCT
		DTC            : UDINT := 16#8B0100;
		DFCid          : UINT  := 101;
		debounceMethod : USINT := TIME_IN_ROW;
	END_STRUCT
END_TYPE
